// TIA Portal project "." (V14)

(* hardware
DEVICE "S7-1200 station_1"  S7-1200 Station
   slot 0: "Rack_0"  S7-1200 Rack  Rack  V1.0
   slot 1: "PLC_1"  CPU 1212C DC/DC/DC  6ES7 212-1AE31-0XB0  V3.0
   slot 2: "AI 4x13BIT/AQ 2x14BIT_1"  SM 1234 AI4/AQ2  6ES7 234-4HE30-0XB0  V1.0
   slot 3: "AI 4xRTD_1"  SM 1231 AI4 x RTD  6ES7 231-5PD32-0XB0  V2.0
   slot 101: "CM 1241 (RS485)_1"  CM 1241 (RS485)  6ES7 241-1CH30-0XB0  V1.0
DEVICE "HMI_1"  KTP600 Basic color PN
   slot 0: "KTP600 Basic color PN"  KTP600 Basic color PN  6AV6 647-0AD11-3AX0  12.0.0.0
   slot 1: "HMI_RT_1"  KTP600 Basic color PN  6AV6 647-0AD11-3AX0  12.0.0.0
   slot 5: "HMI_1.IE_CP_1"  PROFINET Interface  12.0.0.0
      slot 1: "Interfaz PROFINET_1"  PROFINET Interface
         slot 1: "Port_1"  Port
*)

// ===== PLC "PLC_1"  CPU 1212C DC/DC/DC =====

VAR_GLOBAL   // PLC tag table "Tabla de variables estándar"
   "Clock_10Hz" AT %M0.0 : Bool;
   "Clock_5Hz" AT %M0.1 : Bool;
   "Clock_2.5Hz" AT %M0.2 : Bool;
   "Clock_2Hz" AT %M0.3 : Bool;
   "Clock_1.25Hz" AT %M0.4 : Bool;
   "Clock_1Hz" AT %M0.5 : Bool;
   "Clock_0.625Hz" AT %M0.6 : Bool;
   "Clock_0.5Hz" AT %M0.7 : Bool;
   "ConexionExitosa" AT %M5.0 : Bool;
   "AlarmaDesconexion" AT %M5.1 : Bool;
   "A" AT %MW211 : Int;
   "System_Byte" AT %MB1 : Byte;
   "FirstScan" AT %M1.0 : Bool;
   "DiagStatusUpdate" AT %M1.1 : Bool;
   "AlwaysTRUE" AT %M1.2 : Bool;
   "AlwaysFALSE" AT %M1.3 : Bool;
   "ContadorAuxiliar" AT %MW200 : Int;
   "ModoManual" AT %M500.0 : Bool;
   "Tag_1" AT %MD66 : DWord;
   "Tag_2" AT %MD74 : DWord;
END_VAR

VAR_GLOBAL   // PLC tag table "Entradas y Salidas Fisicas"
   "Iniciar" AT %M800.1 : Bool;
   "Extraer" AT %M800.2 : Bool;
   "PilotoVerde" AT %Q0.0 : Bool;
   "PilotoAmarillo" AT %Q0.1 : Bool;
   "PilotoRojo" AT %Q0.2 : Bool;
   "IniciarbOTON" AT %I0.0 : Bool;
   "ExtraerBoton" AT %I0.1 : Bool;
END_VAR

VAR_GLOBAL   // PLC tag table "Memorias de Flanco"
   "Mem_Fer_FlancoBajadaIniciar" AT %M130.1 : Bool;
   "Mem_Fer_FlancoCompleta" AT %M130.2 : Bool;
   "Mem_Des_FlancoDestilado" AT %M131.0 : Bool;
   "Mem_Des_FlancoAgua" AT %M131.2 : Bool;
   "Mem_Rec_FlancoInicio" AT %M132.0 : Bool;
   "Mem_Rec_FlancoObjetivo" AT %M132.1 : Bool;
   "Mem_Rec_FlancoFin" AT %M132.2 : Bool;
   "AlertaAguaBajaDestilador" AT %M132.3 : Bool;
   "NivelBajoDestiador" AT %M132.4 : Bool;
   "Mem_ModoManual_Flanco" AT %M500.1 : Bool;
   "Pulso_SoltarActuadores" AT %M500.2 : Bool;
END_VAR

VAR_GLOBAL   // PLC tag table "Mediciones"
   "Fer_Temperatura" AT %MD40 : Real;
   "Des_Temperatura" AT %MD134 : Real;
   "Fer_Volumen" AT %MD54 : Real;
   "Des_Volumen" AT %MD14 : Real;
   "Rec_Volumen" AT %MD82 : Real;
   "RecirVol" AT %MD92 : Real;
END_VAR

VAR_GLOBAL   // PLC tag table "Estados"
   "Fer_FermentacionCompleta" AT %M72.7 : Bool;
   "Fer_Llenando" AT %M130.0 : Bool;
   "Des_CondicionesClarificar" AT %M131.1 : Bool;
   "AuxAlarmaFermentadorSobrecalentado" AT %MD158 : Real;
END_VAR

VAR_GLOBAL   // PLC tag table "Actuadores"
   "Act_BombaWash" AT %M36.0 : Bool;
   "Act_BombaAguaDestilador" AT %M36.1 : Bool;
   "Act_PurgaDestilador" AT %M36.2 : Bool;
   "Act_ValvRecirculadoDestilador" AT %M36.3 : Bool;
   "Act_ResistenciaDestilador" AT %M36.4 : Bool;
   "Act_ValvIngresoMosto" AT %M72.1 : Bool;
   "Act_PurgaFermentador" AT %M72.2 : Bool;
   "Act_RefrigeracionFermentador" AT %M72.5 : Bool;
   "Act_ValvVaciado" AT %M88.0 : Bool;
   "Act_BombaRecirculado" AT %M90.0 : Bool;
END_VAR

DATA_BLOCK "Proceso"   // DB1
{ S7_Optimized_Access := 'FALSE' }
VERSION : 0.1
   VAR
      Fer_VolInicialMosto : Real := 10.0;
      Fer_LimInfPerdida : Real := 8.12;
      Fer_LimSupTemp : Real := 20.5;
      Fer_LimInfTemp : Real := 19.5;
      Fer_UmbralSobrecalentado : Real := 22.125;
      Des_PesoInicialWash : Real := 0.0;
      Des_AguaAAgregar : Real := 0.0;
      Des_PesoFinal : Real := 0.0;
      Des_VolDescarteMetanol : Real := 0.0;
      Rec_VolBase : Real := 0.0;
      Rec_VolObjetivoRedestilado : Real := 0.0;
   END_VAR
BEGIN
END_DATA_BLOCK

DATA_BLOCK "DatosDeRecetas"   // DB4
{ S7_Optimized_Access := 'FALSE' }
VERSION : 0.1
   VAR
      NombreReceta : String := 'Irlandes';
      NombreReceta_1 : Int := 0;
      SetPointTempFermentador : Real := 20.0;
      HisterisisFermentador : Real := 0.5;
      SetPointTempDestilador : Real := 88.0;
      HisterisisDestilador : Real := 1.0;
      PorcAguaAgregada : Real := 15.0;
      PorcRedestilado : Real := 100.0;
      PorcPerdidaDescarte : Real := 6.125;
      PorcPerdidaFermentacion : Real := 4.0;
      PorcPurgaFermentador : Real := 10.0;
      PorcPurgaDestilador : Real := 5.0;
      CiclosRedestilado : Int := 2;
      VolumenPerdida : Real;
      Fer_LimInfVolumen : Real := 0.125;
      Fer_LimSupVolumen : Real := 52.125;
      Des_LimSupVolumen : Real := 50.125;
      Des_NivelBajo : Real := 0.2;
      Des_LimInfTemp : Real := 87.0;
      Des_LimSupTemp : Real := 89.125;
   END_VAR
BEGIN
END_DATA_BLOCK

DATA_BLOCK "Alarmas"   // DB6
{ S7_Optimized_Access := 'FALSE' }
VERSION : 0.1
   VAR
      Alm_FallaUSS : Bool;
      Alm_FermentadorSobrecalentado : Bool;
      Alm_AvisoDescarteMetanol : Bool;
      Alm_FermentadorLLeno : Bool;
      Alm_DemasiadoWashDestilador : Bool;
      Fase_MomentoDescarteMetanol : Bool;
      Fase_FermentacionTerminada : Bool;
      Fase_InicioLimpiezaFermentador : Bool;
      Fase_FinLimpiezaFermentador : Bool;
      Fase_InicioDestilado : Bool;
      Fase_InicioClarificado : Bool;
      Fase_DescarteExitoso : Bool;
      Fase_WhiskeyTerminado : Bool;
      Fase_InicioRecirculado : Bool;
      Fase_FinRecirculado : Bool;
      Fase_MezclaCompletada : Bool;
      Fase_ContadorRecirculado : Int;
      Vis_FinLimpiezaFermentador : Bool;
      Vis_InicioDestilado : Bool;
      Vis_DescarteExitoso : Bool;
      Vis_AvisoDescarteDeMetanol : Bool;
      aux1 : Bool;
      "aux 2" : Bool;
      AUx : Bool;
      Vis_FinRecirculado : Bool;
      Reserva_HMI : Bool;
   END_VAR
BEGIN
END_DATA_BLOCK

// folder: Control Manual

DATA_BLOCK "ControlManual"   // DB2
{ S7_Optimized_Access := 'FALSE' }
VERSION : 0.1
   VAR
      ManualBombaDeWash : Bool;
      ManualBombaDeAguaDestilador : Bool;
      ManualPurgaDestilador : Bool;
      ManualValvulaRecirculadoDestilador : Bool;
      ManualValvulaIngresoDeMosto : Bool;
      ManualPurgaFermentador : Bool;
      ManualEstadoRefriegeracionFermentador : Bool;
      ManualValvulaDeVaciado : Bool;
      ManualBombaDeRecirculado : Bool;
   END_VAR
BEGIN
END_DATA_BLOCK

// folder: System blocks/Program resources

DATA_BLOCK "IEC_Timer_0_DB"   // DB3
{ S7_Optimized_Access := 'TRUE' }
AUTHOR : Simatic
FAMILY : IEC
NAME : IEC_TMR
VERSION : 1.0
// stored: InstanceOfName IEC_TIMER
"IEC_TIMER"
BEGIN
END_DATA_BLOCK

DATA_BLOCK "IEC_Timer_0_DB_6"   // DB5
{ S7_Optimized_Access := 'TRUE' }
AUTHOR : Simatic
FAMILY : IEC
NAME : IEC_TMR
VERSION : 1.0
// stored: InstanceOfName IEC_TIMER
"IEC_TIMER"
BEGIN
END_DATA_BLOCK

DATA_BLOCK "IEC_Timer_0_DB_7"   // DB7
{ S7_Optimized_Access := 'TRUE' }
AUTHOR : Simatic
FAMILY : IEC
NAME : IEC_TMR
VERSION : 1.0
// stored: InstanceOfName IEC_TIMER
"IEC_TIMER"
BEGIN
END_DATA_BLOCK

DATA_BLOCK "IEC_Timer_0_DB_1"   // DB8
{ S7_Optimized_Access := 'TRUE' }
AUTHOR : Simatic
FAMILY : IEC
NAME : IEC_TMR
VERSION : 1.0
// stored: InstanceOfName IEC_TIMER
"IEC_TIMER"
BEGIN
END_DATA_BLOCK

DATA_BLOCK "IEC_Timer_0_DB_2"   // DB9
{ S7_Optimized_Access := 'TRUE' }
AUTHOR : Simatic
FAMILY : IEC
NAME : IEC_TMR
VERSION : 1.0
// stored: InstanceOfName IEC_TIMER
"IEC_TIMER"
BEGIN
END_DATA_BLOCK

DATA_BLOCK "IEC_Timer_0_DB_3"   // DB10
{ S7_Optimized_Access := 'TRUE' }
AUTHOR : Simatic
FAMILY : IEC
NAME : IEC_TMR
VERSION : 1.0
// stored: InstanceOfName IEC_TIMER
"IEC_TIMER"
BEGIN
END_DATA_BLOCK

DATA_BLOCK "IEC_Timer_0_DB_4"   // DB11
{ S7_Optimized_Access := 'TRUE' }
AUTHOR : Simatic
FAMILY : IEC
NAME : IEC_TMR
VERSION : 1.0
// stored: InstanceOfName IEC_TIMER
"IEC_TIMER"
BEGIN
END_DATA_BLOCK

DATA_BLOCK "IEC_Timer_0_DB_5"   // DB12
{ S7_Optimized_Access := 'TRUE' }
AUTHOR : Simatic
FAMILY : IEC
NAME : IEC_TMR
VERSION : 1.0
// stored: InstanceOfName IEC_TIMER
"IEC_TIMER"
BEGIN
END_DATA_BLOCK

DATA_BLOCK "IEC_Timer_0_DB_9"   // DB13
{ S7_Optimized_Access := 'TRUE' }
AUTHOR : Simatic
FAMILY : IEC
NAME : IEC_TMR
VERSION : 1.0
// stored: InstanceOfName IEC_TIMER
"IEC_TIMER"
BEGIN
END_DATA_BLOCK

DATA_BLOCK "IEC_Timer_0_DB_11"   // DB14
{ S7_Optimized_Access := 'TRUE' }
AUTHOR : Simatic
FAMILY : IEC
NAME : IEC_TMR
VERSION : 1.0
// stored: InstanceOfName IEC_TIMER
"IEC_TIMER"
BEGIN
END_DATA_BLOCK

DATA_BLOCK "IEC_Timer_0_DB_8"   // DB15
{ S7_Optimized_Access := 'TRUE' }
AUTHOR : Simatic
FAMILY : IEC
NAME : IEC_TMR
VERSION : 1.0
// stored: InstanceOfName IEC_TIMER
"IEC_TIMER"
BEGIN
END_DATA_BLOCK

DATA_BLOCK "IEC_Timer_0_DB_10"   // DB17
{ S7_Optimized_Access := 'TRUE' }
AUTHOR : Simatic
FAMILY : IEC
NAME : IEC_TMR
VERSION : 1.0
// stored: InstanceOfName IEC_TIMER
"IEC_TIMER"
BEGIN
END_DATA_BLOCK

// folder: (top level)

ORGANIZATION_BLOCK "control"   // OB126, LAD, ProgramCycle
TITLE = "Main Program Sweep (Cycle)"
{ S7_Optimized_Access := 'TRUE' }
VERSION : 0.1
   VAR_TEMP   // added for the SCL form of the ladder/FBD networks
      _w1 : Bool;
   END_VAR
BEGIN

REGION Network 1
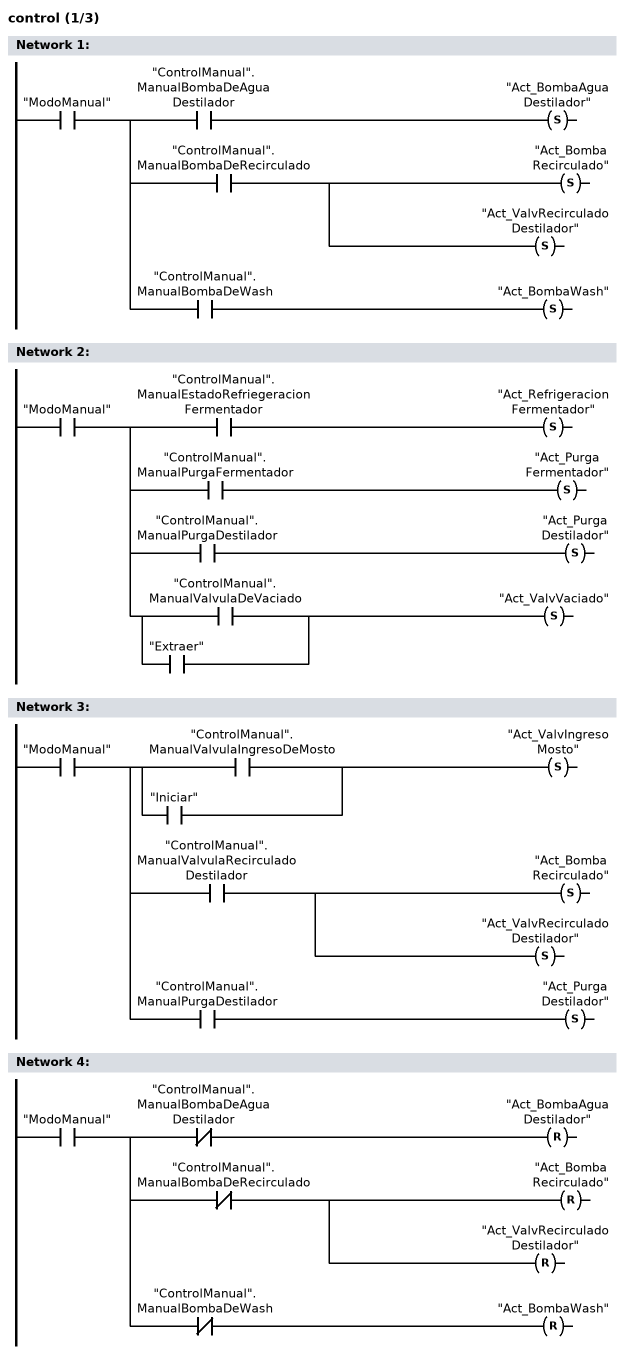
   RUNG wire#powerrail
      Contact( "ModoManual" )
      wire#w1
      Contact( "ControlManual".ManualBombaDeAguaDestilador )
      S_Coil( "Act_BombaAguaDestilador" )
   END_RUNG
   RUNG wire#w1
      Contact( "ControlManual".ManualBombaDeRecirculado )
      wire#w2
      S_Coil( "Act_BombaRecirculado" )
   END_RUNG
   RUNG wire#w2
      S_Coil( "Act_ValvRecirculadoDestilador" )
   END_RUNG
   RUNG wire#w1
      Contact( "ControlManual".ManualBombaDeWash )
      S_Coil( "Act_BombaWash" )
   END_RUNG
   // the same network as SCL:
   IF "ModoManual" AND "ControlManual".ManualBombaDeAguaDestilador THEN
       "Act_BombaAguaDestilador" := TRUE;
   END_IF;
   IF "ModoManual" AND "ControlManual".ManualBombaDeRecirculado THEN
       "Act_BombaRecirculado" := TRUE;
       "Act_ValvRecirculadoDestilador" := TRUE;
   END_IF;
   IF "ModoManual" AND "ControlManual".ManualBombaDeWash THEN "Act_BombaWash" := TRUE; END_IF;
END_REGION

REGION Network 2
   RUNG wire#powerrail
      Contact( "ModoManual" )
      wire#w1
      Contact( "ControlManual".ManualEstadoRefriegeracionFermentador )
      S_Coil( "Act_RefrigeracionFermentador" )
   END_RUNG
   RUNG wire#w1
      Contact( "ControlManual".ManualPurgaFermentador )
      S_Coil( "Act_PurgaFermentador" )
   END_RUNG
   RUNG wire#w1
      Contact( "ControlManual".ManualPurgaDestilador )
      S_Coil( "Act_PurgaDestilador" )
   END_RUNG
   RUNG wire#w1
      Contact( "ControlManual".ManualValvulaDeVaciado )
      wire#w2
      S_Coil( "Act_ValvVaciado" )
   END_RUNG
   RUNG wire#w1
      Contact( "Extraer" )
   END_RUNG wire#w2
   // the same network as SCL:
   IF "ModoManual" AND "ControlManual".ManualEstadoRefriegeracionFermentador THEN
       "Act_RefrigeracionFermentador" := TRUE;
   END_IF;
   IF "ModoManual" AND "ControlManual".ManualPurgaFermentador THEN "Act_PurgaFermentador" := TRUE; END_IF;
   IF "ModoManual" AND "ControlManual".ManualPurgaDestilador THEN "Act_PurgaDestilador" := TRUE; END_IF;
   IF "ModoManual" AND ("ControlManual".ManualValvulaDeVaciado OR "Extraer") THEN
       "Act_ValvVaciado" := TRUE;
   END_IF;
END_REGION

REGION Network 3
   RUNG wire#powerrail
      Contact( "ModoManual" )
      wire#w1
      Contact( "ControlManual".ManualValvulaIngresoDeMosto )
      wire#w2
      S_Coil( "Act_ValvIngresoMosto" )
   END_RUNG
   RUNG wire#w1
      Contact( "Iniciar" )
   END_RUNG wire#w2
   RUNG wire#w1
      Contact( "ControlManual".ManualValvulaRecirculadoDestilador )
      wire#w3
      S_Coil( "Act_BombaRecirculado" )
   END_RUNG
   RUNG wire#w3
      S_Coil( "Act_ValvRecirculadoDestilador" )
   END_RUNG
   RUNG wire#w1
      Contact( "ControlManual".ManualPurgaDestilador )
      S_Coil( "Act_PurgaDestilador" )
   END_RUNG
   // the same network as SCL:
   IF "ModoManual" AND ("ControlManual".ManualValvulaIngresoDeMosto OR "Iniciar") THEN
       "Act_ValvIngresoMosto" := TRUE;
   END_IF;
   IF "ModoManual" AND "ControlManual".ManualValvulaRecirculadoDestilador THEN
       "Act_BombaRecirculado" := TRUE;
       "Act_ValvRecirculadoDestilador" := TRUE;
   END_IF;
   IF "ModoManual" AND "ControlManual".ManualPurgaDestilador THEN "Act_PurgaDestilador" := TRUE; END_IF;
END_REGION

REGION Network 4
   RUNG wire#powerrail
      Contact( "ModoManual" )
      wire#w1
      I_Contact( "ControlManual".ManualBombaDeAguaDestilador )
      R_Coil( "Act_BombaAguaDestilador" )
   END_RUNG
   RUNG wire#w1
      I_Contact( "ControlManual".ManualBombaDeRecirculado )
      wire#w2
      R_Coil( "Act_BombaRecirculado" )
   END_RUNG
   RUNG wire#w2
      R_Coil( "Act_ValvRecirculadoDestilador" )
   END_RUNG
   RUNG wire#w1
      I_Contact( "ControlManual".ManualBombaDeWash )
      R_Coil( "Act_BombaWash" )
   END_RUNG
   // the same network as SCL:
   IF "ModoManual" AND NOT "ControlManual".ManualBombaDeAguaDestilador THEN
       "Act_BombaAguaDestilador" := FALSE;
   END_IF;
   IF "ModoManual" AND NOT "ControlManual".ManualBombaDeRecirculado THEN
       "Act_BombaRecirculado" := FALSE;
       "Act_ValvRecirculadoDestilador" := FALSE;
   END_IF;
   IF "ModoManual" AND NOT "ControlManual".ManualBombaDeWash THEN "Act_BombaWash" := FALSE; END_IF;
END_REGION

REGION Network 5
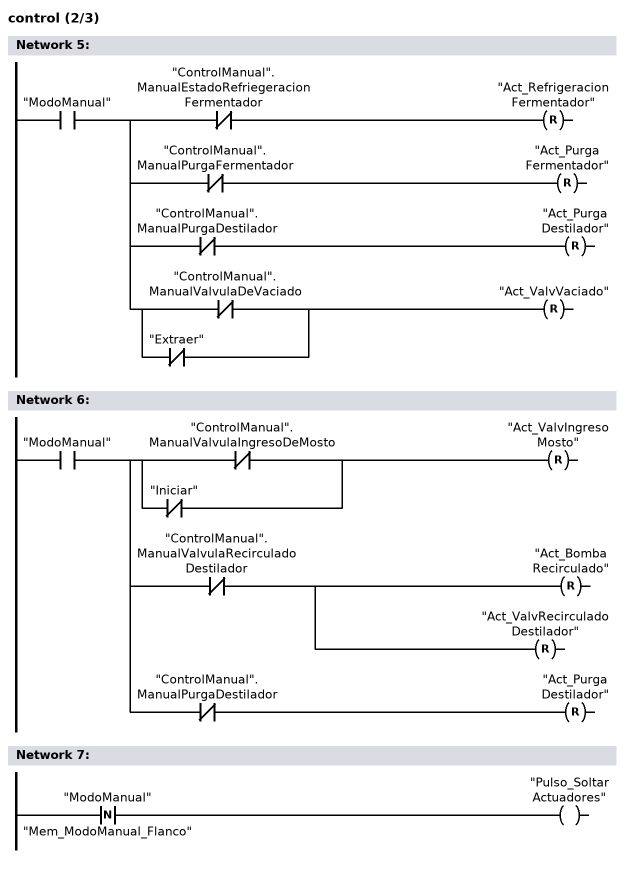
   RUNG wire#powerrail
      Contact( "ModoManual" )
      wire#w1
      I_Contact( "ControlManual".ManualEstadoRefriegeracionFermentador )
      R_Coil( "Act_RefrigeracionFermentador" )
   END_RUNG
   RUNG wire#w1
      I_Contact( "ControlManual".ManualPurgaFermentador )
      R_Coil( "Act_PurgaFermentador" )
   END_RUNG
   RUNG wire#w1
      I_Contact( "ControlManual".ManualPurgaDestilador )
      R_Coil( "Act_PurgaDestilador" )
   END_RUNG
   RUNG wire#w1
      I_Contact( "ControlManual".ManualValvulaDeVaciado )
      wire#w2
      R_Coil( "Act_ValvVaciado" )
   END_RUNG
   RUNG wire#w1
      I_Contact( "Extraer" )
   END_RUNG wire#w2
   // the same network as SCL:
   IF "ModoManual" AND NOT "ControlManual".ManualEstadoRefriegeracionFermentador THEN
       "Act_RefrigeracionFermentador" := FALSE;
   END_IF;
   IF "ModoManual" AND NOT "ControlManual".ManualPurgaFermentador THEN
       "Act_PurgaFermentador" := FALSE;
   END_IF;
   IF "ModoManual" AND NOT "ControlManual".ManualPurgaDestilador THEN "Act_PurgaDestilador" := FALSE; END_IF;
   IF "ModoManual" AND (NOT "ControlManual".ManualValvulaDeVaciado OR NOT "Extraer") THEN
       "Act_ValvVaciado" := FALSE;
   END_IF;
END_REGION

REGION Network 6
   RUNG wire#powerrail
      Contact( "ModoManual" )
      wire#w1
      I_Contact( "ControlManual".ManualValvulaIngresoDeMosto )
      wire#w2
      R_Coil( "Act_ValvIngresoMosto" )
   END_RUNG
   RUNG wire#w1
      I_Contact( "Iniciar" )
   END_RUNG wire#w2
   RUNG wire#w1
      I_Contact( "ControlManual".ManualValvulaRecirculadoDestilador )
      wire#w3
      R_Coil( "Act_BombaRecirculado" )
   END_RUNG
   RUNG wire#w3
      R_Coil( "Act_ValvRecirculadoDestilador" )
   END_RUNG
   RUNG wire#w1
      I_Contact( "ControlManual".ManualPurgaDestilador )
      R_Coil( "Act_PurgaDestilador" )
   END_RUNG
   // the same network as SCL:
   IF "ModoManual" AND (NOT "ControlManual".ManualValvulaIngresoDeMosto OR NOT "Iniciar") THEN
       "Act_ValvIngresoMosto" := FALSE;
   END_IF;
   IF "ModoManual" AND NOT "ControlManual".ManualValvulaRecirculadoDestilador THEN
       "Act_BombaRecirculado" := FALSE;
       "Act_ValvRecirculadoDestilador" := FALSE;
   END_IF;
   IF "ModoManual" AND NOT "ControlManual".ManualPurgaDestilador THEN "Act_PurgaDestilador" := FALSE; END_IF;
END_REGION

REGION Network 7
   RUNG wire#powerrail
      N_Contact(operand := "ModoManual", bit := "Mem_ModoManual_Flanco")
      Coil( "Pulso_SoltarActuadores" )
   END_RUNG
   // the same network as SCL:
   #_w1 := NOT "ModoManual" AND "Mem_ModoManual_Flanco";   // falling edge of "ModoManual"
   "Mem_ModoManual_Flanco" := "ModoManual";
   "Pulso_SoltarActuadores" := #_w1;
END_REGION

REGION Network 8
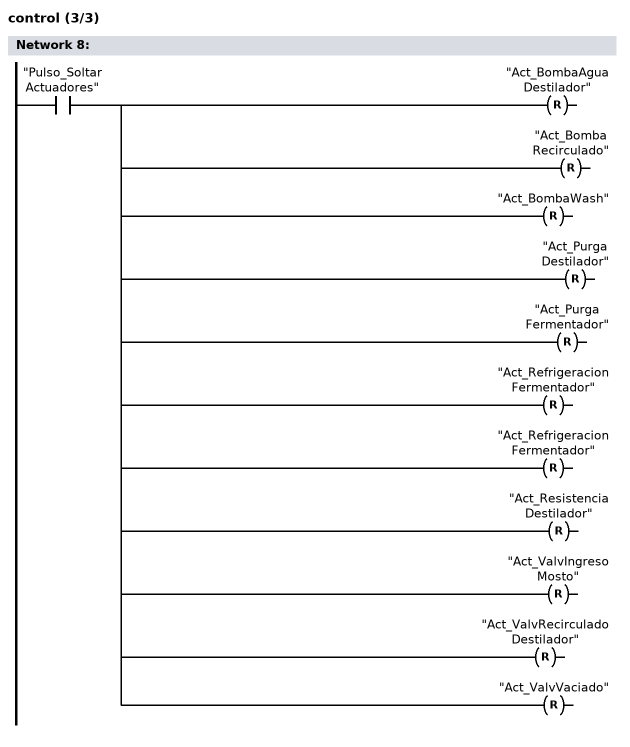
   RUNG wire#powerrail
      Contact( "Pulso_SoltarActuadores" )
      wire#w1
      R_Coil( "Act_BombaAguaDestilador" )
   END_RUNG
   RUNG wire#w1
      R_Coil( "Act_BombaRecirculado" )
   END_RUNG
   RUNG wire#w1
      R_Coil( "Act_BombaWash" )
   END_RUNG
   RUNG wire#w1
      R_Coil( "Act_PurgaDestilador" )
   END_RUNG
   RUNG wire#w1
      R_Coil( "Act_PurgaFermentador" )
   END_RUNG
   RUNG wire#w1
      R_Coil( "Act_RefrigeracionFermentador" )
   END_RUNG
   RUNG wire#w1
      R_Coil( "Act_RefrigeracionFermentador" )
   END_RUNG
   RUNG wire#w1
      R_Coil( "Act_ResistenciaDestilador" )
   END_RUNG
   RUNG wire#w1
      R_Coil( "Act_ValvIngresoMosto" )
   END_RUNG
   RUNG wire#w1
      R_Coil( "Act_ValvRecirculadoDestilador" )
   END_RUNG
   RUNG wire#w1
      R_Coil( "Act_ValvVaciado" )
   END_RUNG
   // the same network as SCL:
   IF "Pulso_SoltarActuadores" THEN
       "Act_BombaAguaDestilador" := FALSE;
       "Act_BombaRecirculado" := FALSE;
       "Act_BombaWash" := FALSE;
       "Act_PurgaDestilador" := FALSE;
       "Act_PurgaFermentador" := FALSE;
       "Act_RefrigeracionFermentador" := FALSE;
       "Act_RefrigeracionFermentador" := FALSE;
       "Act_ResistenciaDestilador" := FALSE;
       "Act_ValvIngresoMosto" := FALSE;
       "Act_ValvRecirculadoDestilador" := FALSE;
       "Act_ValvVaciado" := FALSE;
   END_IF;
END_REGION
END_ORGANIZATION_BLOCK

// folder: Control Manual

ORGANIZATION_BLOCK "Startup"   // OB100, LAD, Startup
TITLE = "Complete Restart"
{ S7_Optimized_Access := 'TRUE' }
VERSION : 0.1
   VAR_INPUT
      LostRetentive : Bool;   // True if retentive data are lost
      LostRTC : Bool;   // True if date and time are lost
   END_VAR
BEGIN

REGION Network 1
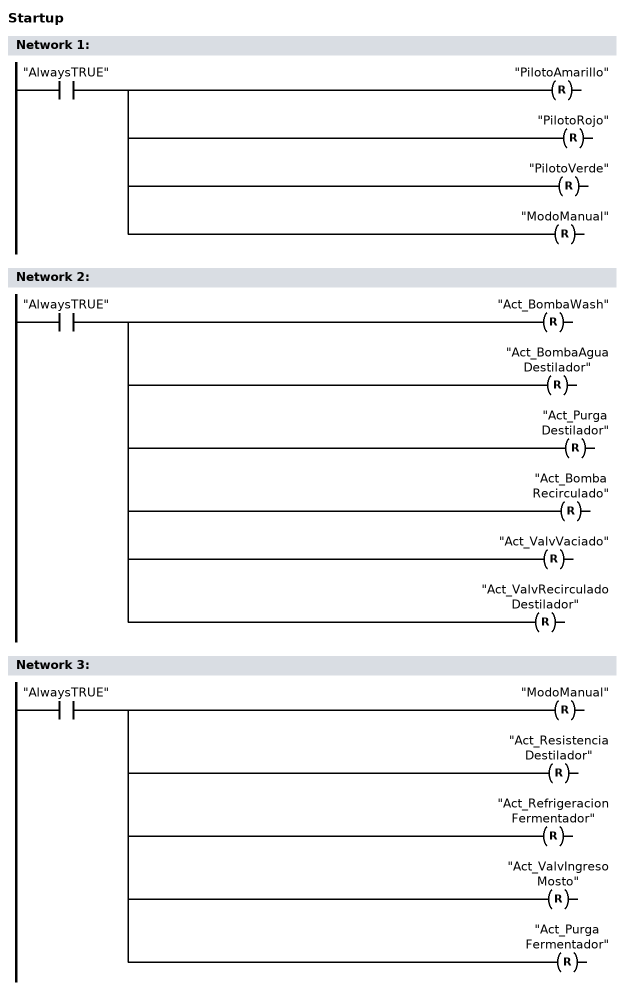
   RUNG wire#powerrail
      Contact( "AlwaysTRUE" )
      wire#w1
      R_Coil( "PilotoAmarillo" )
   END_RUNG
   RUNG wire#w1
      R_Coil( "PilotoRojo" )
   END_RUNG
   RUNG wire#w1
      R_Coil( "PilotoVerde" )
   END_RUNG
   RUNG wire#w1
      R_Coil( "ModoManual" )
   END_RUNG
   // the same network as SCL:
   IF "AlwaysTRUE" THEN
       "PilotoAmarillo" := FALSE;
       "PilotoRojo" := FALSE;
       "PilotoVerde" := FALSE;
       "ModoManual" := FALSE;
   END_IF;
END_REGION

REGION Network 2
   RUNG wire#powerrail
      Contact( "AlwaysTRUE" )
      wire#w1
      R_Coil( "Act_BombaWash" )
   END_RUNG
   RUNG wire#w1
      R_Coil( "Act_BombaAguaDestilador" )
   END_RUNG
   RUNG wire#w1
      R_Coil( "Act_PurgaDestilador" )
   END_RUNG
   RUNG wire#w1
      R_Coil( "Act_BombaRecirculado" )
   END_RUNG
   RUNG wire#w1
      R_Coil( "Act_ValvVaciado" )
   END_RUNG
   RUNG wire#w1
      R_Coil( "Act_ValvRecirculadoDestilador" )
   END_RUNG
   // the same network as SCL:
   IF "AlwaysTRUE" THEN
       "Act_BombaWash" := FALSE;
       "Act_BombaAguaDestilador" := FALSE;
       "Act_PurgaDestilador" := FALSE;
       "Act_BombaRecirculado" := FALSE;
       "Act_ValvVaciado" := FALSE;
       "Act_ValvRecirculadoDestilador" := FALSE;
   END_IF;
END_REGION

REGION Network 3
   RUNG wire#powerrail
      Contact( "AlwaysTRUE" )
      wire#w1
      R_Coil( "ModoManual" )
   END_RUNG
   RUNG wire#w1
      R_Coil( "Act_ResistenciaDestilador" )
   END_RUNG
   RUNG wire#w1
      R_Coil( "Act_RefrigeracionFermentador" )
   END_RUNG
   RUNG wire#w1
      R_Coil( "Act_ValvIngresoMosto" )
   END_RUNG
   RUNG wire#w1
      R_Coil( "Act_PurgaFermentador" )
   END_RUNG
   // the same network as SCL:
   IF "AlwaysTRUE" THEN
       "ModoManual" := FALSE;
       "Act_ResistenciaDestilador" := FALSE;
       "Act_RefrigeracionFermentador" := FALSE;
       "Act_ValvIngresoMosto" := FALSE;
       "Act_PurgaFermentador" := FALSE;
   END_IF;
END_REGION
END_ORGANIZATION_BLOCK

// folder: Destilador

ORGANIZATION_BLOCK "Control de Temperatura destilador"   // OB31, LAD, CyclicInterrupt
{ S7_Optimized_Access := 'TRUE' }
VERSION : 0.1
   VAR_TEMP   // added for the SCL form of the ladder/FBD networks
      _w1 : Bool;
      _w2 : Bool;
   END_VAR
BEGIN

REGION Network 1: Control
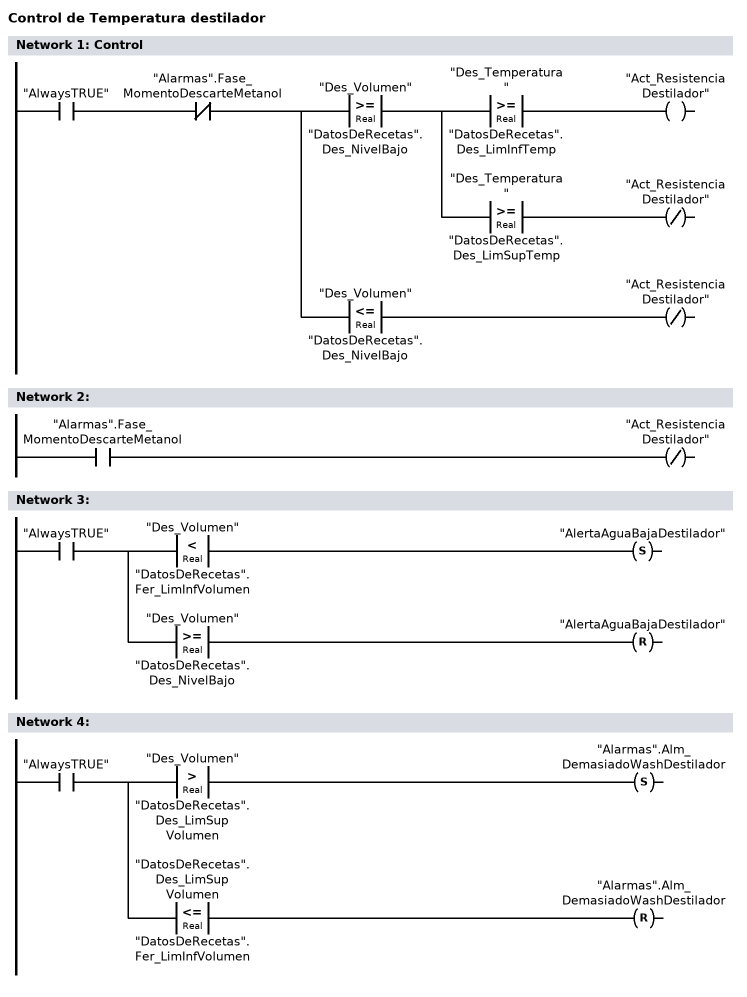
   RUNG wire#powerrail
      Contact( "AlwaysTRUE" )
      I_Contact( "Alarmas".Fase_MomentoDescarteMetanol )
      wire#w1
      { S7_Templates := "SrcType := Real" } GE_Contact(in1 := "Des_Volumen", in2 := "DatosDeRecetas".Des_NivelBajo)
      wire#w2
      { S7_Templates := "SrcType := Real" } GE_Contact(in1 := "Des_Temperatura", in2 := "DatosDeRecetas".Des_LimInfTemp)
      Coil( "Act_ResistenciaDestilador" )
   END_RUNG
   RUNG wire#w2
      { S7_Templates := "SrcType := Real" } GE_Contact(in1 := "Des_Temperatura", in2 := "DatosDeRecetas".Des_LimSupTemp)
      I_Coil( "Act_ResistenciaDestilador" )
   END_RUNG
   RUNG wire#w1
      { S7_Templates := "SrcType := Real" } LE_Contact(in1 := "Des_Volumen", in2 := "DatosDeRecetas".Des_NivelBajo)
      I_Coil( "Act_ResistenciaDestilador" )
   END_RUNG
   // the same network as SCL:
   #_w1 := "AlwaysTRUE" AND NOT "Alarmas".Fase_MomentoDescarteMetanol;
   #_w2 := #_w1 AND ("Des_Volumen" >= "DatosDeRecetas".Des_NivelBajo);
   "Act_ResistenciaDestilador" := #_w2 AND ("Des_Temperatura" >= "DatosDeRecetas".Des_LimInfTemp);
   "Act_ResistenciaDestilador" := NOT (#_w2 AND ("Des_Temperatura" >= "DatosDeRecetas".Des_LimSupTemp));
   "Act_ResistenciaDestilador" := NOT (#_w1 AND ("Des_Volumen" <= "DatosDeRecetas".Des_NivelBajo));
END_REGION

REGION Network 2
   RUNG wire#powerrail
      Contact( "Alarmas".Fase_MomentoDescarteMetanol )
      I_Coil( "Act_ResistenciaDestilador" )
   END_RUNG
   // the same network as SCL:
   "Act_ResistenciaDestilador" := NOT "Alarmas".Fase_MomentoDescarteMetanol;
END_REGION

REGION Network 3
   RUNG wire#powerrail
      Contact( "AlwaysTRUE" )
      wire#w1
      { S7_Templates := "SrcType := Real" } LT_Contact(in1 := "Des_Volumen", in2 := "DatosDeRecetas".Fer_LimInfVolumen)
      S_Coil( "AlertaAguaBajaDestilador" )
   END_RUNG
   RUNG wire#w1
      { S7_Templates := "SrcType := Real" } GE_Contact(in1 := "Des_Volumen", in2 := "DatosDeRecetas".Des_NivelBajo)
      R_Coil( "AlertaAguaBajaDestilador" )
   END_RUNG
   // the same network as SCL:
   IF "AlwaysTRUE" AND ("Des_Volumen" < "DatosDeRecetas".Fer_LimInfVolumen) THEN
       "AlertaAguaBajaDestilador" := TRUE;
   END_IF;
   IF "AlwaysTRUE" AND ("Des_Volumen" >= "DatosDeRecetas".Des_NivelBajo) THEN
       "AlertaAguaBajaDestilador" := FALSE;
   END_IF;
END_REGION

REGION Network 4
   RUNG wire#powerrail
      Contact( "AlwaysTRUE" )
      wire#w1
      { S7_Templates := "SrcType := Real" } GT_Contact(in1 := "Des_Volumen", in2 := "DatosDeRecetas".Des_LimSupVolumen)
      S_Coil( "Alarmas".Alm_DemasiadoWashDestilador )
   END_RUNG
   RUNG wire#w1
      { S7_Templates := "SrcType := Real" } LE_Contact(in1 := "DatosDeRecetas".Des_LimSupVolumen, in2 := "DatosDeRecetas".Fer_LimInfVolumen)
      R_Coil( "Alarmas".Alm_DemasiadoWashDestilador )
   END_RUNG
   // the same network as SCL:
   IF "AlwaysTRUE" AND ("Des_Volumen" > "DatosDeRecetas".Des_LimSupVolumen) THEN
       "Alarmas".Alm_DemasiadoWashDestilador := TRUE;
   END_IF;
   IF "AlwaysTRUE" AND ("DatosDeRecetas".Des_LimSupVolumen <= "DatosDeRecetas".Fer_LimInfVolumen) THEN
       "Alarmas".Alm_DemasiadoWashDestilador := FALSE;
   END_IF;
END_REGION
END_ORGANIZATION_BLOCK

ORGANIZATION_BLOCK "Configuracion y ciclo de programa"   // OB124, LAD, ProgramCycle
TITLE = "Main Program Sweep (Cycle)"
{ S7_Optimized_Access := 'TRUE' }
VERSION : 0.1
   VAR_TEMP
      PesoInicialDelWash : Real;
      Temp_1 : Bool;
      PesoFinal : Real;
      AguaAAgregar : Real;
      PesoDeMetanol : Real;
   END_VAR
   VAR_TEMP   // added for the SCL form of the ladder/FBD networks
      _w1 : Bool;
   END_VAR
BEGIN

REGION Network 1: Pesaje previo al clarificado
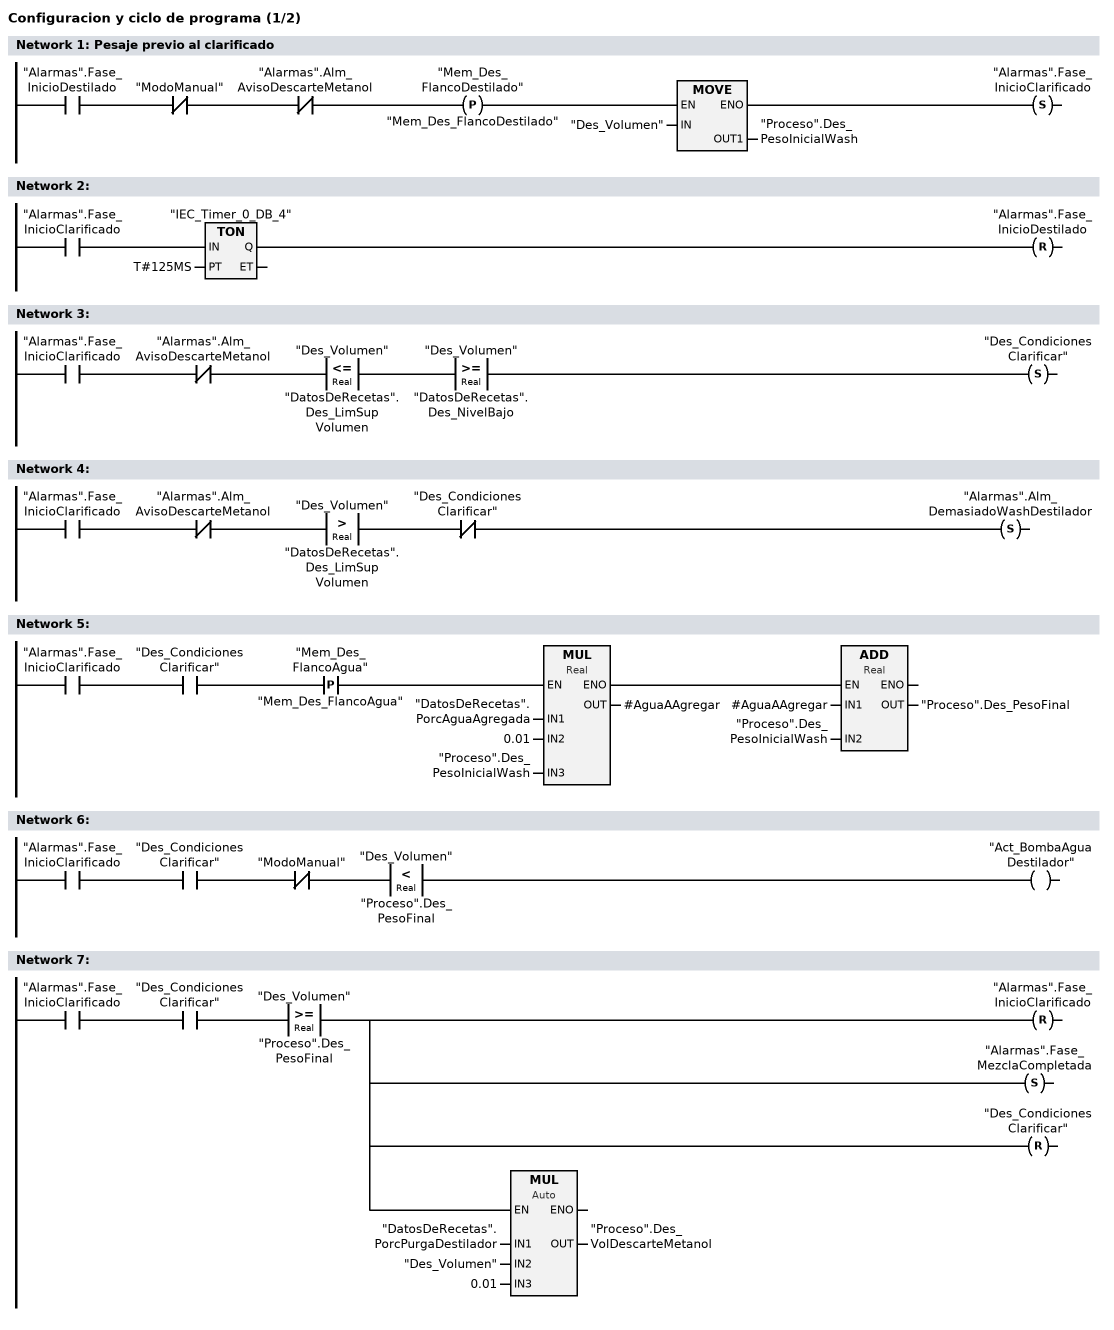
   // ENO of a box is taken as its EN; it also drops when the box reports an error
   #_w1 := "Alarmas".Fase_InicioDestilado AND NOT "ModoManual" AND NOT "Alarmas".Alm_AvisoDescarteMetanol;
   "Mem_Des_FlancoDestilado" := #_w1 AND NOT "Mem_Des_FlancoDestilado";   // rising edge
   "Mem_Des_FlancoDestilado" := #_w1;
   IF #_w1 THEN
       "Proceso".Des_PesoInicialWash := "Des_Volumen";
       "Alarmas".Fase_InicioClarificado := TRUE;
   END_IF;
END_REGION

REGION Network 2
   "IEC_Timer_0_DB_4".TON(IN := "Alarmas".Fase_InicioClarificado, PT := T#125MS);
   IF "IEC_Timer_0_DB_4".Q THEN "Alarmas".Fase_InicioDestilado := FALSE; END_IF;
END_REGION

REGION Network 3
   RUNG wire#powerrail
      Contact( "Alarmas".Fase_InicioClarificado )
      I_Contact( "Alarmas".Alm_AvisoDescarteMetanol )
      { S7_Templates := "SrcType := Real" } LE_Contact(in1 := "Des_Volumen", in2 := "DatosDeRecetas".Des_LimSupVolumen)
      { S7_Templates := "SrcType := Real" } GE_Contact(in1 := "Des_Volumen", in2 := "DatosDeRecetas".Des_NivelBajo)
      S_Coil( "Des_CondicionesClarificar" )
   END_RUNG
   // the same network as SCL:
   IF "Alarmas".Fase_InicioClarificado AND NOT "Alarmas".Alm_AvisoDescarteMetanol AND ("Des_Volumen" <= "DatosDeRecetas".Des_LimSupVolumen) AND ("Des_Volumen" >= "DatosDeRecetas".Des_NivelBajo) THEN
       "Des_CondicionesClarificar" := TRUE;
   END_IF;
END_REGION

REGION Network 4
   RUNG wire#powerrail
      Contact( "Alarmas".Fase_InicioClarificado )
      I_Contact( "Alarmas".Alm_AvisoDescarteMetanol )
      { S7_Templates := "SrcType := Real" } GT_Contact(in1 := "Des_Volumen", in2 := "DatosDeRecetas".Des_LimSupVolumen)
      I_Contact( "Des_CondicionesClarificar" )
      S_Coil( "Alarmas".Alm_DemasiadoWashDestilador )
   END_RUNG
   // the same network as SCL:
   IF "Alarmas".Fase_InicioClarificado AND NOT "Alarmas".Alm_AvisoDescarteMetanol AND ("Des_Volumen" > "DatosDeRecetas".Des_LimSupVolumen) AND NOT "Des_CondicionesClarificar" THEN
       "Alarmas".Alm_DemasiadoWashDestilador := TRUE;
   END_IF;
END_REGION

REGION Network 5
   RUNG wire#powerrail
      Contact( "Alarmas".Fase_InicioClarificado )
      Contact( "Des_CondicionesClarificar" )
      P_Contact(operand := "Mem_Des_FlancoAgua", bit := "Mem_Des_FlancoAgua")
      { S7_Templates := "SrcType := Real"; S7_GenerateENO := "TRUE" } Mul(in1 := "DatosDeRecetas".PorcAguaAgregada, in2 := 0.01, in3 := "Proceso".Des_PesoInicialWash, out => #AguaAAgregar)
      { S7_Templates := "SrcType := Real"; S7_GenerateENO := "TRUE" } Add(in1 := #AguaAAgregar, in2 := "Proceso".Des_PesoInicialWash, out => "Proceso".Des_PesoFinal)
   END_RUNG
   // the same network as SCL:
   // ENO of a box is taken as its EN; it also drops when the box reports an error
   #_w1 := "Alarmas".Fase_InicioClarificado AND "Des_CondicionesClarificar" AND "Mem_Des_FlancoAgua" AND NOT "Mem_Des_FlancoAgua";   // rising edge of "Mem_Des_FlancoAgua"
   "Mem_Des_FlancoAgua" := "Mem_Des_FlancoAgua";
   IF #_w1 THEN
       #AguaAAgregar := "DatosDeRecetas".PorcAguaAgregada * 0.01 * "Proceso".Des_PesoInicialWash;
       "Proceso".Des_PesoFinal := #AguaAAgregar + "Proceso".Des_PesoInicialWash;
   END_IF;
END_REGION

REGION Network 6
   RUNG wire#powerrail
      Contact( "Alarmas".Fase_InicioClarificado )
      Contact( "Des_CondicionesClarificar" )
      I_Contact( "ModoManual" )
      { S7_Templates := "SrcType := Real" } LT_Contact(in1 := "Des_Volumen", in2 := "Proceso".Des_PesoFinal)
      Coil( "Act_BombaAguaDestilador" )
   END_RUNG
   // the same network as SCL:
   "Act_BombaAguaDestilador" := "Alarmas".Fase_InicioClarificado AND "Des_CondicionesClarificar" AND NOT "ModoManual" AND ("Des_Volumen" < "Proceso".Des_PesoFinal);
END_REGION

REGION Network 7
   RUNG wire#powerrail
      Contact( "Alarmas".Fase_InicioClarificado )
      Contact( "Des_CondicionesClarificar" )
      { S7_Templates := "SrcType := Real" } GE_Contact(in1 := "Des_Volumen", in2 := "Proceso".Des_PesoFinal)
      wire#w1
      R_Coil( "Alarmas".Fase_InicioClarificado )
   END_RUNG
   RUNG wire#w1
      S_Coil( "Alarmas".Fase_MezclaCompletada )
   END_RUNG
   RUNG wire#w1
      R_Coil( "Des_CondicionesClarificar" )
   END_RUNG
   RUNG wire#w1
      { S7_GenerateENO := "TRUE" } Mul(in1 := "DatosDeRecetas".PorcPurgaDestilador, in2 := "Des_Volumen", in3 := 0.01, out => "Proceso".Des_VolDescarteMetanol)
   END_RUNG
   // the same network as SCL:
   #_w1 := "Alarmas".Fase_InicioClarificado AND "Des_CondicionesClarificar" AND ("Des_Volumen" >= "Proceso".Des_PesoFinal);
   IF #_w1 THEN
       "Alarmas".Fase_InicioClarificado := FALSE;
       "Alarmas".Fase_MezclaCompletada := TRUE;
       "Des_CondicionesClarificar" := FALSE;
       "Proceso".Des_VolDescarteMetanol := "DatosDeRecetas".PorcPurgaDestilador * "Des_Volumen" * 0.01;
   END_IF;
END_REGION

REGION Network 8
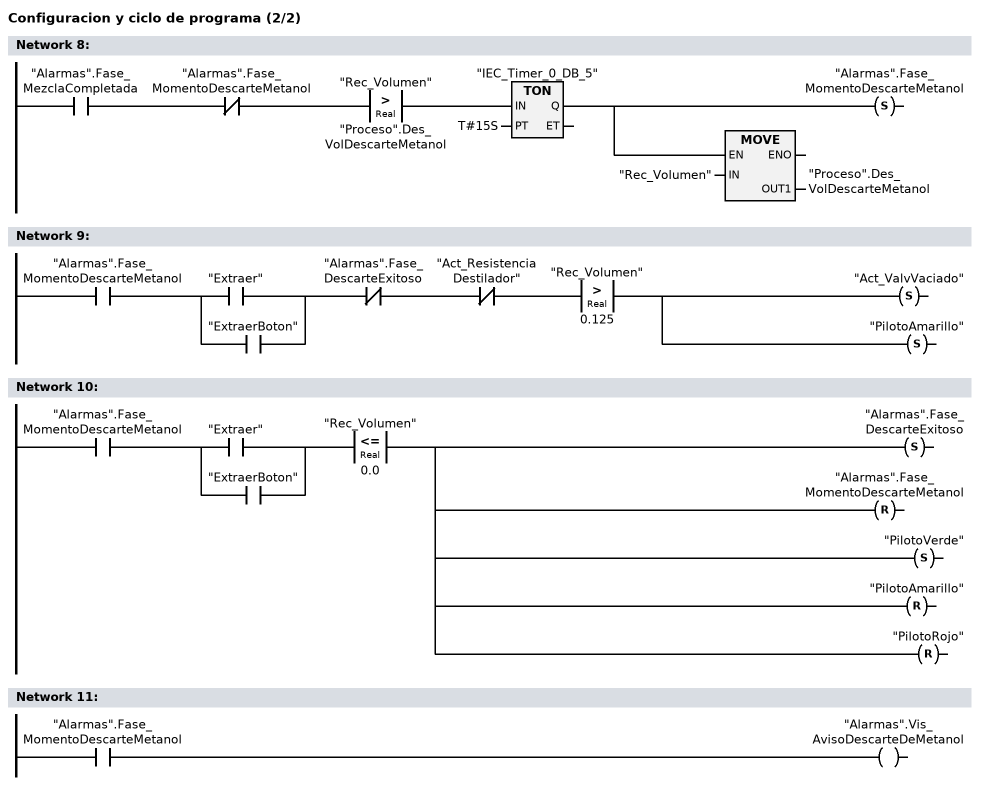
   "IEC_Timer_0_DB_5".TON(IN := "Alarmas".Fase_MezclaCompletada AND NOT "Alarmas".Fase_MomentoDescarteMetanol AND ("Rec_Volumen" > "Proceso".Des_VolDescarteMetanol),
                          PT := T#15S);
   IF "IEC_Timer_0_DB_5".Q THEN
       "Alarmas".Fase_MomentoDescarteMetanol := TRUE;
       "Proceso".Des_VolDescarteMetanol := "Rec_Volumen";
   END_IF;
END_REGION

REGION Network 9
   RUNG wire#powerrail
      Contact( "Alarmas".Fase_MomentoDescarteMetanol )
      wire#w1
      Contact( "Extraer" )
      wire#w2
      I_Contact( "Alarmas".Fase_DescarteExitoso )
      I_Contact( "Act_ResistenciaDestilador" )
      { S7_Templates := "SrcType := Real" } GT_Contact(in1 := "Rec_Volumen", in2 := 0.125)
      wire#w3
      S_Coil( "Act_ValvVaciado" )
   END_RUNG
   RUNG wire#w1
      Contact( "ExtraerBoton" )
   END_RUNG wire#w2
   RUNG wire#w3
      S_Coil( "PilotoAmarillo" )
   END_RUNG
   // the same network as SCL:
   IF "Alarmas".Fase_MomentoDescarteMetanol AND ("Extraer" OR "ExtraerBoton") AND NOT "Alarmas".Fase_DescarteExitoso AND NOT "Act_ResistenciaDestilador" AND ("Rec_Volumen" > 0.125) THEN
       "Act_ValvVaciado" := TRUE;
       "PilotoAmarillo" := TRUE;
   END_IF;
END_REGION

REGION Network 10
   RUNG wire#powerrail
      Contact( "Alarmas".Fase_MomentoDescarteMetanol )
      wire#w1
      Contact( "Extraer" )
      wire#w2
      { S7_Templates := "SrcType := Real" } LE_Contact(in1 := "Rec_Volumen", in2 := 0.0)
      wire#w3
      S_Coil( "Alarmas".Fase_DescarteExitoso )
   END_RUNG
   RUNG wire#w1
      Contact( "ExtraerBoton" )
   END_RUNG wire#w2
   RUNG wire#w3
      R_Coil( "Alarmas".Fase_MomentoDescarteMetanol )
   END_RUNG
   RUNG wire#w3
      S_Coil( "PilotoVerde" )
   END_RUNG
   RUNG wire#w3
      R_Coil( "PilotoAmarillo" )
   END_RUNG
   RUNG wire#w3
      R_Coil( "PilotoRojo" )
   END_RUNG
   // the same network as SCL:
   IF "Alarmas".Fase_MomentoDescarteMetanol AND ("Extraer" OR "ExtraerBoton") AND ("Rec_Volumen" <= 0.0) THEN
       "Alarmas".Fase_DescarteExitoso := TRUE;
   END_IF;
   #_w1 := "Alarmas".Fase_MomentoDescarteMetanol AND ("Extraer" OR "ExtraerBoton") AND ("Rec_Volumen" <= 0.0);
   IF #_w1 THEN
       "Alarmas".Fase_MomentoDescarteMetanol := FALSE;
       "PilotoVerde" := TRUE;
       "PilotoAmarillo" := FALSE;
       "PilotoRojo" := FALSE;
   END_IF;
END_REGION

REGION Network 11
   RUNG wire#powerrail
      Contact( "Alarmas".Fase_MomentoDescarteMetanol )
      Coil( "Alarmas".Vis_AvisoDescarteDeMetanol )
   END_RUNG
   // the same network as SCL:
   "Alarmas".Vis_AvisoDescarteDeMetanol := "Alarmas".Fase_MomentoDescarteMetanol;
END_REGION
END_ORGANIZATION_BLOCK

ORGANIZATION_BLOCK "Calcular  limites on off destilador"   // OB127, LAD, ProgramCycle
TITLE = "Main Program Sweep (Cycle)"
{ S7_Optimized_Access := 'TRUE' }
VERSION : 0.1
BEGIN

REGION Network 1
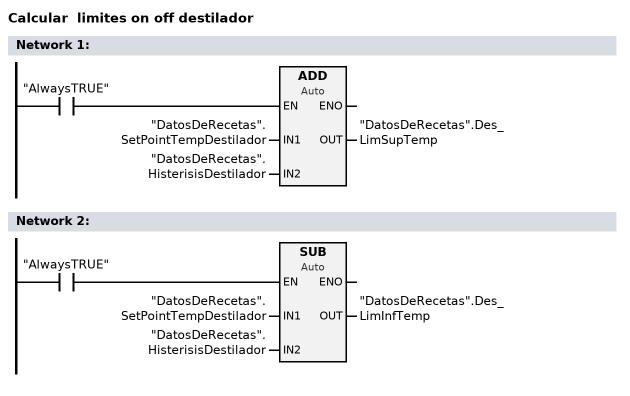
   RUNG wire#powerrail
      Contact( "AlwaysTRUE" )
      { S7_GenerateENO := "TRUE" } Add(in1 := "DatosDeRecetas".SetPointTempDestilador, in2 := "DatosDeRecetas".HisterisisDestilador, out => "DatosDeRecetas".Des_LimSupTemp)
   END_RUNG
   // the same network as SCL:
   IF "AlwaysTRUE" THEN
       "DatosDeRecetas".Des_LimSupTemp := "DatosDeRecetas".SetPointTempDestilador + "DatosDeRecetas".HisterisisDestilador;
   END_IF;
END_REGION

REGION Network 2
   RUNG wire#powerrail
      Contact( "AlwaysTRUE" )
      { S7_GenerateENO := "TRUE" } Sub(in1 := "DatosDeRecetas".SetPointTempDestilador, in2 := "DatosDeRecetas".HisterisisDestilador, out => "DatosDeRecetas".Des_LimInfTemp)
   END_RUNG
   // the same network as SCL:
   IF "AlwaysTRUE" THEN
       "DatosDeRecetas".Des_LimInfTemp := "DatosDeRecetas".SetPointTempDestilador - "DatosDeRecetas".HisterisisDestilador;
   END_IF;
END_REGION
END_ORGANIZATION_BLOCK

// folder: Fermentador

ORGANIZATION_BLOCK "Control de ingreso Mosto y salida de Wash"   // OB1, LAD, ProgramCycle
TITLE = "Control del Mosto y Wash Fermentador"
{ S7_Optimized_Access := 'TRUE' }
VERSION : 0.1
   VAR_TEMP
      Auxiliarrr : Real;
      FlancoDeBajadaInicio : Bool;
      Temp_1 : Bool;
      Auxiliar : Bool;
   END_VAR
   VAR_TEMP   // added for the SCL form of the ladder/FBD networks
      _w1 : Bool;
   END_VAR
BEGIN

REGION Network 1
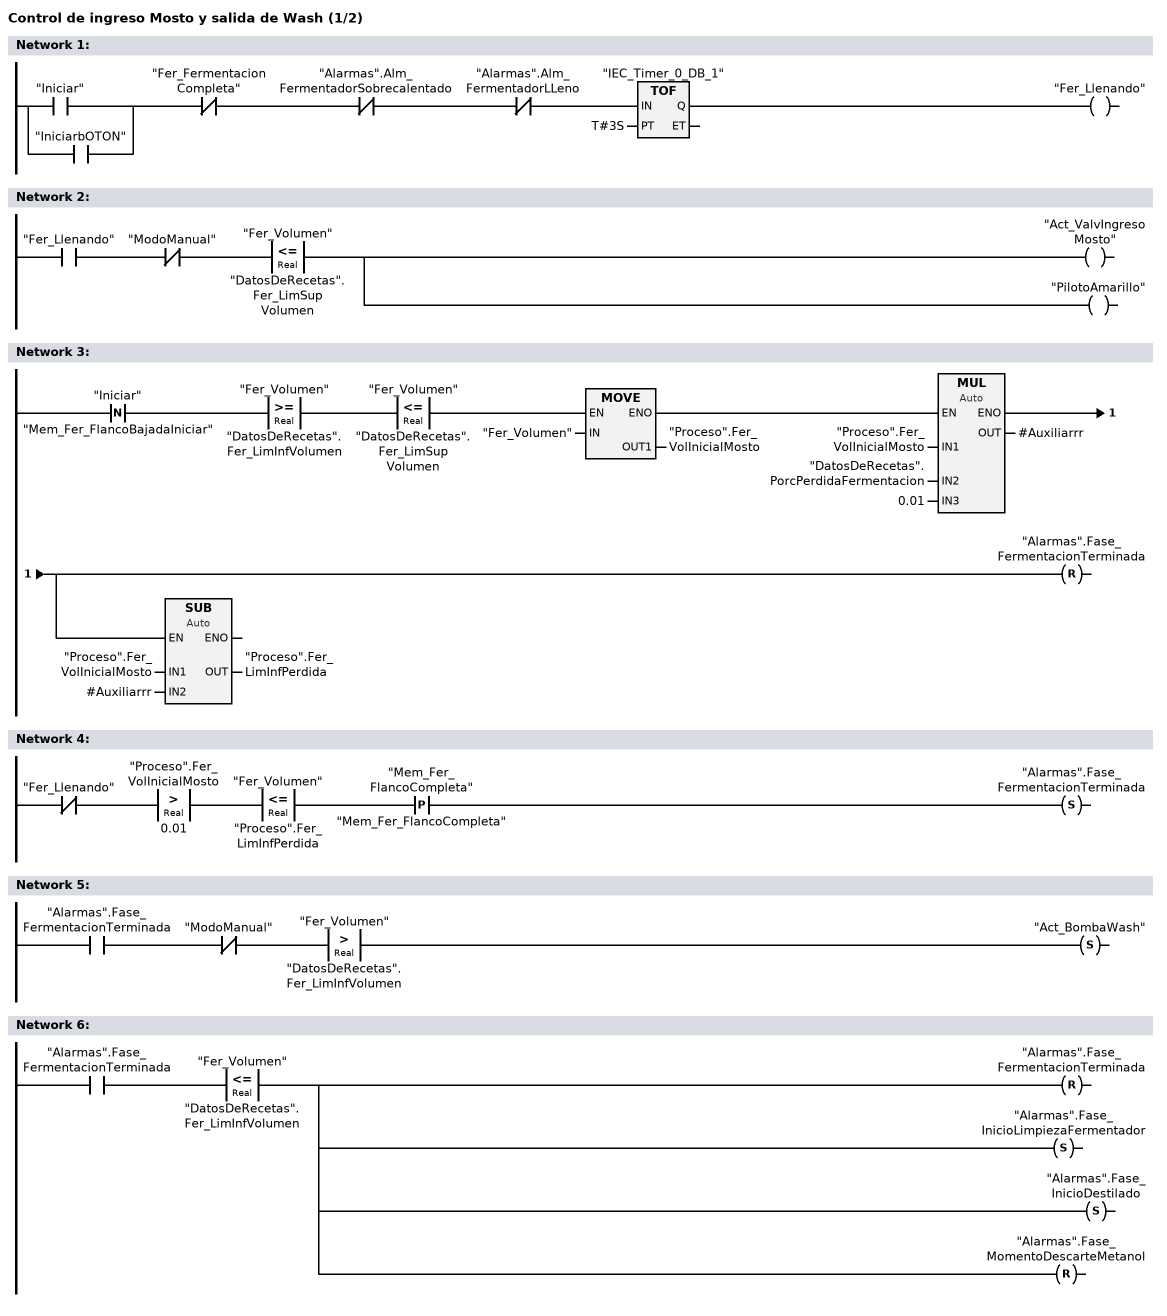
   "IEC_Timer_0_DB_1".TOF(IN := ("Iniciar" OR "IniciarbOTON") AND NOT "Fer_FermentacionCompleta" AND NOT "Alarmas".Alm_FermentadorSobrecalentado AND NOT "Alarmas".Alm_FermentadorLLeno,
                          PT := T#3S);
   "Fer_Llenando" := "IEC_Timer_0_DB_1".Q;
END_REGION

REGION Network 2
   RUNG wire#powerrail
      Contact( "Fer_Llenando" )
      I_Contact( "ModoManual" )
      { S7_Templates := "SrcType := Real" } LE_Contact(in1 := "Fer_Volumen", in2 := "DatosDeRecetas".Fer_LimSupVolumen)
      wire#w1
      Coil( "Act_ValvIngresoMosto" )
   END_RUNG
   RUNG wire#w1
      Coil( "PilotoAmarillo" )
   END_RUNG
   // the same network as SCL:
   "Act_ValvIngresoMosto" := "Fer_Llenando" AND NOT "ModoManual" AND ("Fer_Volumen" <= "DatosDeRecetas".Fer_LimSupVolumen);
   "PilotoAmarillo" := "Act_ValvIngresoMosto";
END_REGION

REGION Network 3
   RUNG wire#powerrail
      N_Contact(operand := "Iniciar", bit := "Mem_Fer_FlancoBajadaIniciar")
      { S7_Templates := "SrcType := Real" } GE_Contact(in1 := "Fer_Volumen", in2 := "DatosDeRecetas".Fer_LimInfVolumen)
      { S7_Templates := "SrcType := Real" } LE_Contact(in1 := "Fer_Volumen", in2 := "DatosDeRecetas".Fer_LimSupVolumen)
      { S7_GenerateENO := "TRUE" } Move(in := "Fer_Volumen", out1 => "Proceso".Fer_VolInicialMosto)
      { S7_GenerateENO := "TRUE" } Mul(in1 := "Proceso".Fer_VolInicialMosto, in2 := "DatosDeRecetas".PorcPerdidaFermentacion, in3 := 0.01, out => #Auxiliarrr)
      wire#w1
      R_Coil( "Alarmas".Fase_FermentacionTerminada )
   END_RUNG
   RUNG wire#w1
      { S7_GenerateENO := "TRUE" } Sub(in1 := "Proceso".Fer_VolInicialMosto, in2 := #Auxiliarrr, out => "Proceso".Fer_LimInfPerdida)
   END_RUNG
   // the same network as SCL:
   // ENO of a box is taken as its EN; it also drops when the box reports an error
   #_w1 := NOT "Iniciar" AND "Mem_Fer_FlancoBajadaIniciar";   // falling edge of "Iniciar"
   "Mem_Fer_FlancoBajadaIniciar" := "Iniciar";
   IF #_w1 AND ("Fer_Volumen" >= "DatosDeRecetas".Fer_LimInfVolumen) AND ("Fer_Volumen" <= "DatosDeRecetas".Fer_LimSupVolumen) THEN
       "Proceso".Fer_VolInicialMosto := "Fer_Volumen";
       #Auxiliarrr := "Proceso".Fer_VolInicialMosto * "DatosDeRecetas".PorcPerdidaFermentacion * 0.01;
       "Alarmas".Fase_FermentacionTerminada := FALSE;
       "Proceso".Fer_LimInfPerdida := "Proceso".Fer_VolInicialMosto - #Auxiliarrr;
   END_IF;
END_REGION

REGION Network 4
   RUNG wire#powerrail
      I_Contact( "Fer_Llenando" )
      { S7_Templates := "SrcType := Real" } GT_Contact(in1 := "Proceso".Fer_VolInicialMosto, in2 := 0.01)
      { S7_Templates := "SrcType := Real" } LE_Contact(in1 := "Fer_Volumen", in2 := "Proceso".Fer_LimInfPerdida)
      P_Contact(operand := "Mem_Fer_FlancoCompleta", bit := "Mem_Fer_FlancoCompleta")
      S_Coil( "Alarmas".Fase_FermentacionTerminada )
   END_RUNG
   // the same network as SCL:
   #_w1 := NOT "Fer_Llenando" AND ("Proceso".Fer_VolInicialMosto > 0.01) AND ("Fer_Volumen" <= "Proceso".Fer_LimInfPerdida) AND "Mem_Fer_FlancoCompleta" AND NOT "Mem_Fer_FlancoCompleta";   // rising edge of "Mem_Fer_FlancoCompleta"
   "Mem_Fer_FlancoCompleta" := "Mem_Fer_FlancoCompleta";
   IF #_w1 THEN "Alarmas".Fase_FermentacionTerminada := TRUE; END_IF;
END_REGION

REGION Network 5
   RUNG wire#powerrail
      Contact( "Alarmas".Fase_FermentacionTerminada )
      I_Contact( "ModoManual" )
      { S7_Templates := "SrcType := Real" } GT_Contact(in1 := "Fer_Volumen", in2 := "DatosDeRecetas".Fer_LimInfVolumen)
      S_Coil( "Act_BombaWash" )
   END_RUNG
   // the same network as SCL:
   IF "Alarmas".Fase_FermentacionTerminada AND NOT "ModoManual" AND ("Fer_Volumen" > "DatosDeRecetas".Fer_LimInfVolumen) THEN
       "Act_BombaWash" := TRUE;
   END_IF;
END_REGION

REGION Network 6
   RUNG wire#powerrail
      Contact( "Alarmas".Fase_FermentacionTerminada )
      { S7_Templates := "SrcType := Real" } LE_Contact(in1 := "Fer_Volumen", in2 := "DatosDeRecetas".Fer_LimInfVolumen)
      wire#w1
      R_Coil( "Alarmas".Fase_FermentacionTerminada )
   END_RUNG
   RUNG wire#w1
      S_Coil( "Alarmas".Fase_InicioLimpiezaFermentador )
   END_RUNG
   RUNG wire#w1
      S_Coil( "Alarmas".Fase_InicioDestilado )
   END_RUNG
   RUNG wire#w1
      R_Coil( "Alarmas".Fase_MomentoDescarteMetanol )
   END_RUNG
   // the same network as SCL:
   #_w1 := "Alarmas".Fase_FermentacionTerminada AND ("Fer_Volumen" <= "DatosDeRecetas".Fer_LimInfVolumen);
   IF #_w1 THEN
       "Alarmas".Fase_FermentacionTerminada := FALSE;
       "Alarmas".Fase_InicioLimpiezaFermentador := TRUE;
       "Alarmas".Fase_InicioDestilado := TRUE;
       "Alarmas".Fase_MomentoDescarteMetanol := FALSE;
   END_IF;
END_REGION

REGION Network 7
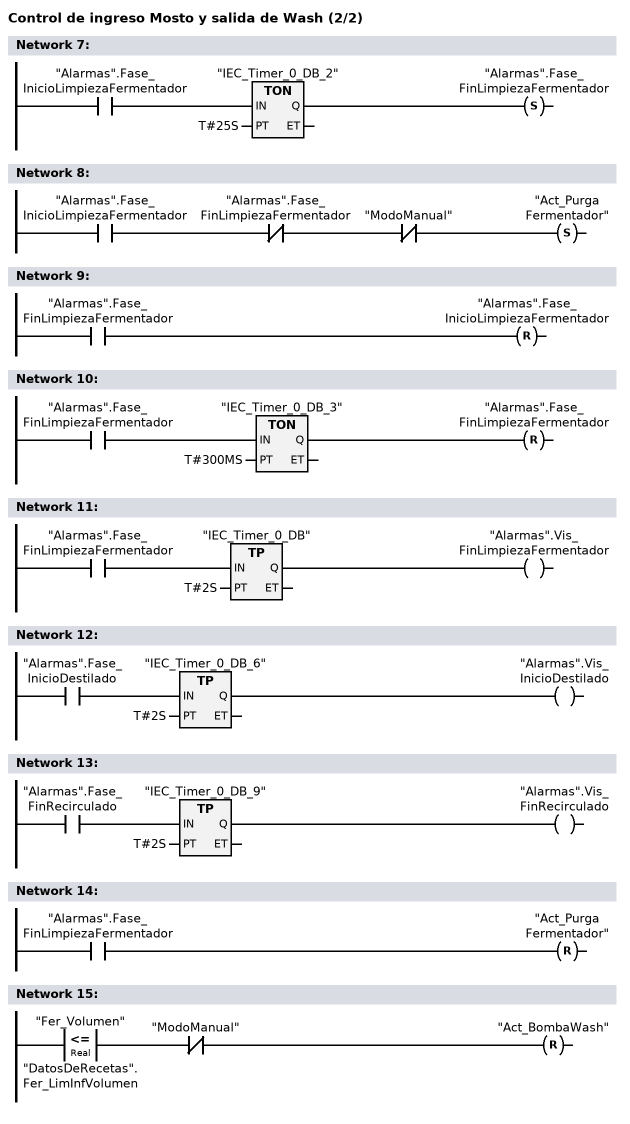
   "IEC_Timer_0_DB_2".TON(IN := "Alarmas".Fase_InicioLimpiezaFermentador, PT := T#25S);
   IF "IEC_Timer_0_DB_2".Q THEN "Alarmas".Fase_FinLimpiezaFermentador := TRUE; END_IF;
END_REGION

REGION Network 8
   RUNG wire#powerrail
      Contact( "Alarmas".Fase_InicioLimpiezaFermentador )
      I_Contact( "Alarmas".Fase_FinLimpiezaFermentador )
      I_Contact( "ModoManual" )
      S_Coil( "Act_PurgaFermentador" )
   END_RUNG
   // the same network as SCL:
   IF "Alarmas".Fase_InicioLimpiezaFermentador AND NOT "Alarmas".Fase_FinLimpiezaFermentador AND NOT "ModoManual" THEN
       "Act_PurgaFermentador" := TRUE;
   END_IF;
END_REGION

REGION Network 9
   RUNG wire#powerrail
      Contact( "Alarmas".Fase_FinLimpiezaFermentador )
      R_Coil( "Alarmas".Fase_InicioLimpiezaFermentador )
   END_RUNG
   // the same network as SCL:
   IF "Alarmas".Fase_FinLimpiezaFermentador THEN "Alarmas".Fase_InicioLimpiezaFermentador := FALSE; END_IF;
END_REGION

REGION Network 10
   "IEC_Timer_0_DB_3".TON(IN := "Alarmas".Fase_FinLimpiezaFermentador, PT := T#300MS);
   IF "IEC_Timer_0_DB_3".Q THEN "Alarmas".Fase_FinLimpiezaFermentador := FALSE; END_IF;
END_REGION

REGION Network 11
   "IEC_Timer_0_DB".TP(IN := "Alarmas".Fase_FinLimpiezaFermentador, PT := T#2S);
   "Alarmas".Vis_FinLimpiezaFermentador := "IEC_Timer_0_DB".Q;
END_REGION

REGION Network 12
   "IEC_Timer_0_DB_6".TP(IN := "Alarmas".Fase_InicioDestilado, PT := T#2S);
   "Alarmas".Vis_InicioDestilado := "IEC_Timer_0_DB_6".Q;
END_REGION

REGION Network 13
   "IEC_Timer_0_DB_9".TP(IN := "Alarmas".Fase_FinRecirculado, PT := T#2S);
   "Alarmas".Vis_FinRecirculado := "IEC_Timer_0_DB_9".Q;
END_REGION

REGION Network 14
   RUNG wire#powerrail
      Contact( "Alarmas".Fase_FinLimpiezaFermentador )
      R_Coil( "Act_PurgaFermentador" )
   END_RUNG
   // the same network as SCL:
   IF "Alarmas".Fase_FinLimpiezaFermentador THEN "Act_PurgaFermentador" := FALSE; END_IF;
END_REGION

REGION Network 15
   RUNG wire#powerrail
      { S7_Templates := "SrcType := Real" } LE_Contact(in1 := "Fer_Volumen", in2 := "DatosDeRecetas".Fer_LimInfVolumen)
      I_Contact( "ModoManual" )
      R_Coil( "Act_BombaWash" )
   END_RUNG
   // the same network as SCL:
   IF ("Fer_Volumen" <= "DatosDeRecetas".Fer_LimInfVolumen) AND NOT "ModoManual" THEN
       "Act_BombaWash" := FALSE;
   END_IF;
END_REGION
END_ORGANIZATION_BLOCK

ORGANIZATION_BLOCK "Control De Temperatura Del Fermentador"   // OB123, LAD, ProgramCycle
TITLE = "Main Program Sweep (Cycle)" / Control e la temperatura del Fermentador
{ S7_Optimized_Access := 'TRUE' }
VERSION : 0.1
// Nuestro fermentador solo tiene banda negativa; no tiene resistencia calefactora, solo refrigeración, esto tiene una razon de ser, al tratarse de una planta  en una zona cálida no se corre riesgo de que las levaduras mueran por el frío, si de calor y se avinagre el wash
   VAR_TEMP
      LimiteInferiorTemperatura : Real;
      LimiteSuperiorTemperatura : Real;
   END_VAR
   VAR_TEMP   // added for the SCL form of the ladder/FBD networks
      _w1 : Bool;
   END_VAR
BEGIN

REGION Network 1
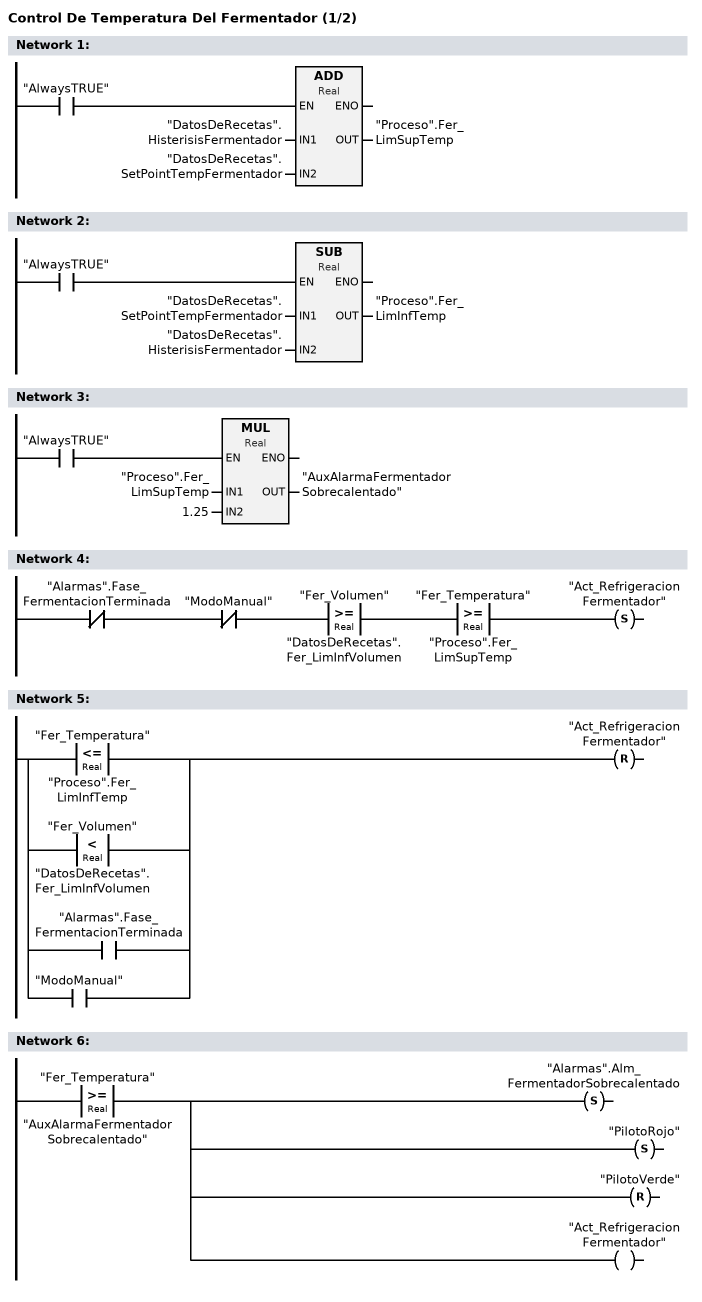
   RUNG wire#powerrail
      Contact( "AlwaysTRUE" )
      { S7_Templates := "SrcType := Real"; S7_GenerateENO := "TRUE" } Add(in1 := "DatosDeRecetas".HisterisisFermentador, in2 := "DatosDeRecetas".SetPointTempFermentador, out => "Proceso".Fer_LimSupTemp)
   END_RUNG
   // the same network as SCL:
   IF "AlwaysTRUE" THEN
       "Proceso".Fer_LimSupTemp := "DatosDeRecetas".HisterisisFermentador + "DatosDeRecetas".SetPointTempFermentador;
   END_IF;
END_REGION

REGION Network 2
   RUNG wire#powerrail
      Contact( "AlwaysTRUE" )
      { S7_Templates := "SrcType := Real"; S7_GenerateENO := "TRUE" } Sub(in1 := "DatosDeRecetas".SetPointTempFermentador, in2 := "DatosDeRecetas".HisterisisFermentador, out => "Proceso".Fer_LimInfTemp)
   END_RUNG
   // the same network as SCL:
   IF "AlwaysTRUE" THEN
       "Proceso".Fer_LimInfTemp := "DatosDeRecetas".SetPointTempFermentador - "DatosDeRecetas".HisterisisFermentador;
   END_IF;
END_REGION

REGION Network 3
   RUNG wire#powerrail
      Contact( "AlwaysTRUE" )
      { S7_Templates := "SrcType := Real"; S7_GenerateENO := "TRUE" } Mul(in1 := "Proceso".Fer_LimSupTemp, in2 := 1.25, out => "AuxAlarmaFermentadorSobrecalentado")
   END_RUNG
   // the same network as SCL:
   IF "AlwaysTRUE" THEN "AuxAlarmaFermentadorSobrecalentado" := "Proceso".Fer_LimSupTemp * 1.25; END_IF;
END_REGION

REGION Network 4
   RUNG wire#powerrail
      I_Contact( "Alarmas".Fase_FermentacionTerminada )
      I_Contact( "ModoManual" )
      { S7_Templates := "SrcType := Real" } GE_Contact(in1 := "Fer_Volumen", in2 := "DatosDeRecetas".Fer_LimInfVolumen)
      { S7_Templates := "SrcType := Real" } GE_Contact(in1 := "Fer_Temperatura", in2 := "Proceso".Fer_LimSupTemp)
      S_Coil( "Act_RefrigeracionFermentador" )
   END_RUNG
   // the same network as SCL:
   IF NOT "Alarmas".Fase_FermentacionTerminada AND NOT "ModoManual" AND ("Fer_Volumen" >= "DatosDeRecetas".Fer_LimInfVolumen) AND ("Fer_Temperatura" >= "Proceso".Fer_LimSupTemp) THEN
       "Act_RefrigeracionFermentador" := TRUE;
   END_IF;
END_REGION

REGION Network 5
   RUNG wire#powerrail
      { S7_Templates := "SrcType := Real" } LE_Contact(in1 := "Fer_Temperatura", in2 := "Proceso".Fer_LimInfTemp)
      wire#w1
      R_Coil( "Act_RefrigeracionFermentador" )
   END_RUNG
   RUNG wire#powerrail
      { S7_Templates := "SrcType := Real" } LT_Contact(in1 := "Fer_Volumen", in2 := "DatosDeRecetas".Fer_LimInfVolumen)
   END_RUNG wire#w1
   RUNG wire#powerrail
      Contact( "Alarmas".Fase_FermentacionTerminada )
   END_RUNG wire#w1
   RUNG wire#powerrail
      Contact( "ModoManual" )
   END_RUNG wire#w1
   // the same network as SCL:
   IF ("Fer_Temperatura" <= "Proceso".Fer_LimInfTemp) OR ("Fer_Volumen" < "DatosDeRecetas".Fer_LimInfVolumen) OR "Alarmas".Fase_FermentacionTerminada OR "ModoManual" THEN
       "Act_RefrigeracionFermentador" := FALSE;
   END_IF;
END_REGION

REGION Network 6
   RUNG wire#powerrail
      { S7_Templates := "SrcType := Real" } GE_Contact(in1 := "Fer_Temperatura", in2 := "AuxAlarmaFermentadorSobrecalentado")
      wire#w1
      S_Coil( "Alarmas".Alm_FermentadorSobrecalentado )
   END_RUNG
   RUNG wire#w1
      S_Coil( "PilotoRojo" )
   END_RUNG
   RUNG wire#w1
      R_Coil( "PilotoVerde" )
   END_RUNG
   RUNG wire#w1
      Coil( "Act_RefrigeracionFermentador" )
   END_RUNG
   // the same network as SCL:
   #_w1 := "Fer_Temperatura" >= "AuxAlarmaFermentadorSobrecalentado";
   IF #_w1 THEN
       "Alarmas".Alm_FermentadorSobrecalentado := TRUE;
       "PilotoRojo" := TRUE;
       "PilotoVerde" := FALSE;
   END_IF;
   "Act_RefrigeracionFermentador" := #_w1;
END_REGION

REGION Network 7
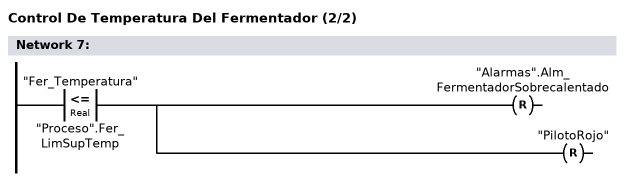
   RUNG wire#powerrail
      { S7_Templates := "SrcType := Real" } LE_Contact(in1 := "Fer_Temperatura", in2 := "Proceso".Fer_LimSupTemp)
      wire#w1
      R_Coil( "Alarmas".Alm_FermentadorSobrecalentado )
   END_RUNG
   RUNG wire#w1
      R_Coil( "PilotoRojo" )
   END_RUNG
   // the same network as SCL:
   IF "Fer_Temperatura" <= "Proceso".Fer_LimSupTemp THEN
       "Alarmas".Alm_FermentadorSobrecalentado := FALSE;
       "PilotoRojo" := FALSE;
   END_IF;
END_REGION
END_ORGANIZATION_BLOCK

// folder: Tanques

ORGANIZATION_BLOCK "Recirculado"   // OB125, LAD, ProgramCycle
TITLE = "Main Program Sweep (Cycle)"
{ S7_Optimized_Access := 'TRUE' }
VERSION : 0.1
   VAR_TEMP
      Impulso : Bool;
      InicioImpulso : Bool;
      Auxiliar : Real;
   END_VAR
   VAR CONSTANT
      Uno : Int := 1;
   END_VAR
   VAR_TEMP   // added for the SCL form of the ladder/FBD networks
      _w1 : Bool;
   END_VAR
BEGIN

REGION Network 1
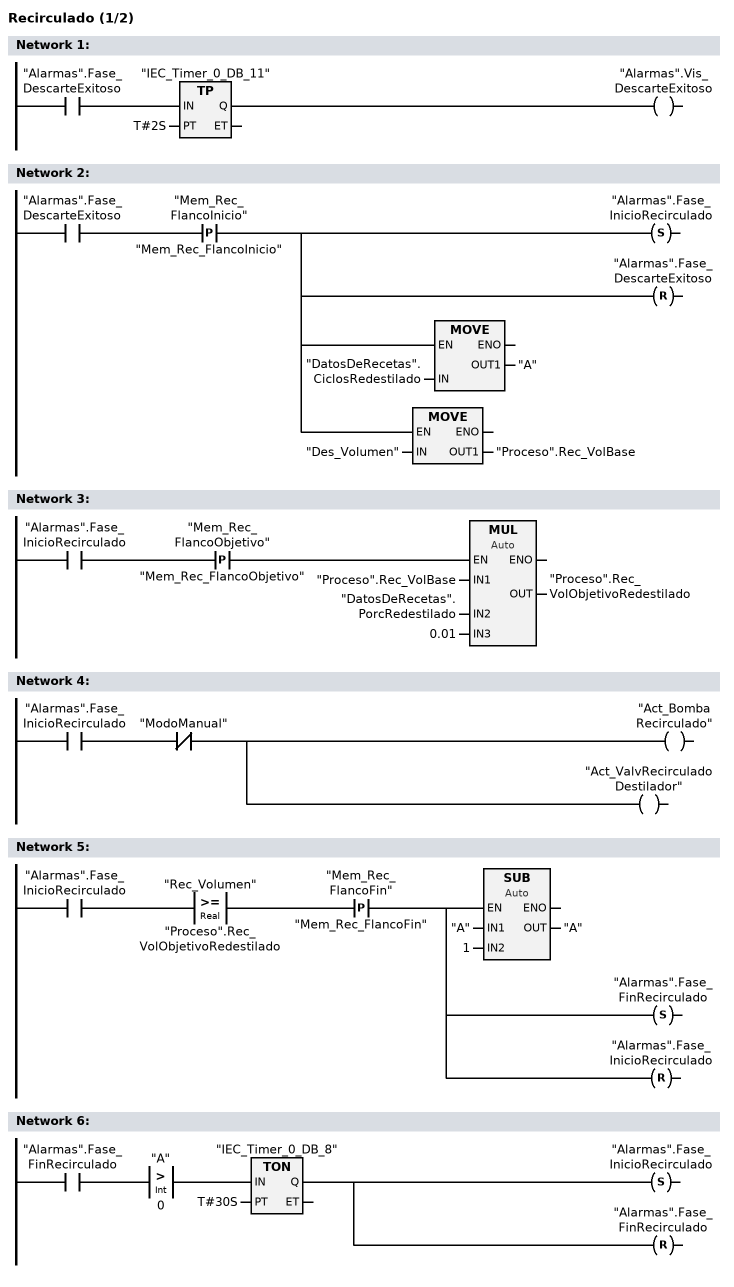
   "IEC_Timer_0_DB_11".TP(IN := "Alarmas".Fase_DescarteExitoso, PT := T#2S);
   "Alarmas".Vis_DescarteExitoso := "IEC_Timer_0_DB_11".Q;
END_REGION

REGION Network 2
   RUNG wire#powerrail
      Contact( "Alarmas".Fase_DescarteExitoso )
      P_Contact(operand := "Mem_Rec_FlancoInicio", bit := "Mem_Rec_FlancoInicio")
      wire#w1
      S_Coil( "Alarmas".Fase_InicioRecirculado )
   END_RUNG
   RUNG wire#w1
      R_Coil( "Alarmas".Fase_DescarteExitoso )
   END_RUNG
   RUNG wire#w1
      { S7_GenerateENO := "TRUE" } Move(in := "DatosDeRecetas".CiclosRedestilado, out1 => "A")
   END_RUNG
   RUNG wire#w1
      { S7_GenerateENO := "TRUE" } Move(in := "Des_Volumen", out1 => "Proceso".Rec_VolBase)
   END_RUNG
   // the same network as SCL:
   #_w1 := "Alarmas".Fase_DescarteExitoso AND "Mem_Rec_FlancoInicio" AND NOT "Mem_Rec_FlancoInicio";   // rising edge of "Mem_Rec_FlancoInicio"
   "Mem_Rec_FlancoInicio" := "Mem_Rec_FlancoInicio";
   IF #_w1 THEN
       "Alarmas".Fase_InicioRecirculado := TRUE;
       "Alarmas".Fase_DescarteExitoso := FALSE;
       "A" := "DatosDeRecetas".CiclosRedestilado;
       "Proceso".Rec_VolBase := "Des_Volumen";
   END_IF;
END_REGION

REGION Network 3
   RUNG wire#powerrail
      Contact( "Alarmas".Fase_InicioRecirculado )
      P_Contact(operand := "Mem_Rec_FlancoObjetivo", bit := "Mem_Rec_FlancoObjetivo")
      { S7_GenerateENO := "TRUE" } Mul(in1 := "Proceso".Rec_VolBase, in2 := "DatosDeRecetas".PorcRedestilado, in3 := 0.01, out => "Proceso".Rec_VolObjetivoRedestilado)
   END_RUNG
   // the same network as SCL:
   #_w1 := "Alarmas".Fase_InicioRecirculado AND "Mem_Rec_FlancoObjetivo" AND NOT "Mem_Rec_FlancoObjetivo";   // rising edge of "Mem_Rec_FlancoObjetivo"
   "Mem_Rec_FlancoObjetivo" := "Mem_Rec_FlancoObjetivo";
   IF #_w1 THEN
       "Proceso".Rec_VolObjetivoRedestilado := "Proceso".Rec_VolBase * "DatosDeRecetas".PorcRedestilado * 0.01;
   END_IF;
END_REGION

REGION Network 4
   RUNG wire#powerrail
      Contact( "Alarmas".Fase_InicioRecirculado )
      I_Contact( "ModoManual" )
      wire#w1
      Coil( "Act_BombaRecirculado" )
   END_RUNG
   RUNG wire#w1
      Coil( "Act_ValvRecirculadoDestilador" )
   END_RUNG
   // the same network as SCL:
   "Act_BombaRecirculado" := "Alarmas".Fase_InicioRecirculado AND NOT "ModoManual";
   "Act_ValvRecirculadoDestilador" := "Act_BombaRecirculado";
END_REGION

REGION Network 5
   RUNG wire#powerrail
      Contact( "Alarmas".Fase_InicioRecirculado )
      { S7_Templates := "SrcType := Real" } GE_Contact(in1 := "Rec_Volumen", in2 := "Proceso".Rec_VolObjetivoRedestilado)
      P_Contact(operand := "Mem_Rec_FlancoFin", bit := "Mem_Rec_FlancoFin")
      wire#w1
      { S7_GenerateENO := "TRUE" } Sub(in1 := "A", in2 := 1, out => "A")
   END_RUNG
   RUNG wire#w1
      S_Coil( "Alarmas".Fase_FinRecirculado )
   END_RUNG
   RUNG wire#w1
      R_Coil( "Alarmas".Fase_InicioRecirculado )
   END_RUNG
   // the same network as SCL:
   #_w1 := "Alarmas".Fase_InicioRecirculado AND ("Rec_Volumen" >= "Proceso".Rec_VolObjetivoRedestilado) AND "Mem_Rec_FlancoFin" AND NOT "Mem_Rec_FlancoFin";   // rising edge of "Mem_Rec_FlancoFin"
   "Mem_Rec_FlancoFin" := "Mem_Rec_FlancoFin";
   IF #_w1 THEN
       "A" := "A" - 1;
       "Alarmas".Fase_FinRecirculado := TRUE;
       "Alarmas".Fase_InicioRecirculado := FALSE;
   END_IF;
END_REGION

REGION Network 6
   "IEC_Timer_0_DB_8".TON(IN := "Alarmas".Fase_FinRecirculado AND ("A" > 0), PT := T#30S);
   IF "IEC_Timer_0_DB_8".Q THEN
       "Alarmas".Fase_InicioRecirculado := TRUE;
       "Alarmas".Fase_FinRecirculado := FALSE;
   END_IF;
END_REGION

REGION Network 7
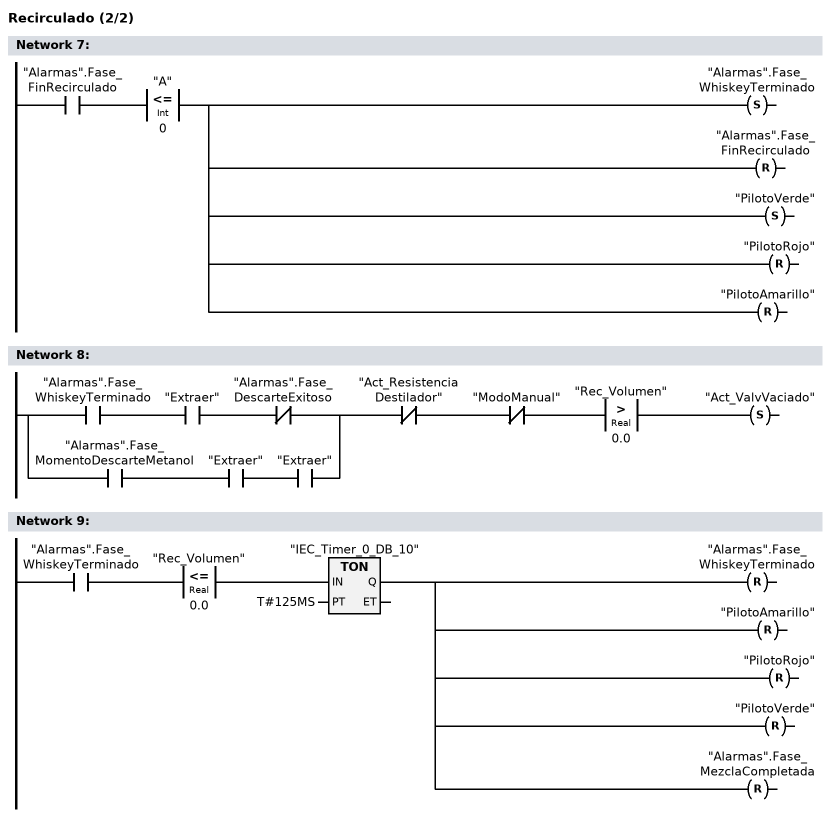
   RUNG wire#powerrail
      Contact( "Alarmas".Fase_FinRecirculado )
      { S7_Templates := "SrcType := Int" } LE_Contact(in1 := "A", in2 := 0)
      wire#w1
      S_Coil( "Alarmas".Fase_WhiskeyTerminado )
   END_RUNG
   RUNG wire#w1
      R_Coil( "Alarmas".Fase_FinRecirculado )
   END_RUNG
   RUNG wire#w1
      S_Coil( "PilotoVerde" )
   END_RUNG
   RUNG wire#w1
      R_Coil( "PilotoRojo" )
   END_RUNG
   RUNG wire#w1
      R_Coil( "PilotoAmarillo" )
   END_RUNG
   // the same network as SCL:
   IF "Alarmas".Fase_FinRecirculado AND ("A" <= 0) THEN "Alarmas".Fase_WhiskeyTerminado := TRUE; END_IF;
   #_w1 := "Alarmas".Fase_FinRecirculado AND ("A" <= 0);
   IF #_w1 THEN
       "Alarmas".Fase_FinRecirculado := FALSE;
       "PilotoVerde" := TRUE;
       "PilotoRojo" := FALSE;
       "PilotoAmarillo" := FALSE;
   END_IF;
END_REGION

REGION Network 8
   RUNG wire#powerrail
      Contact( "Alarmas".Fase_WhiskeyTerminado )
      Contact( "Extraer" )
      I_Contact( "Alarmas".Fase_DescarteExitoso )
      wire#w1
      I_Contact( "Act_ResistenciaDestilador" )
      I_Contact( "ModoManual" )
      { S7_Templates := "SrcType := Real" } GT_Contact(in1 := "Rec_Volumen", in2 := 0.0)
      S_Coil( "Act_ValvVaciado" )
   END_RUNG
   RUNG wire#powerrail
      Contact( "Alarmas".Fase_MomentoDescarteMetanol )
      Contact( "Extraer" )
      Contact( "Extraer" )
   END_RUNG wire#w1
   // the same network as SCL:
   IF (("Alarmas".Fase_WhiskeyTerminado AND "Extraer" AND NOT "Alarmas".Fase_DescarteExitoso) OR ("Alarmas".Fase_MomentoDescarteMetanol AND "Extraer" AND "Extraer")) AND NOT "Act_ResistenciaDestilador" AND NOT "ModoManual" AND ("Rec_Volumen" > 0.0) THEN
       "Act_ValvVaciado" := TRUE;
   END_IF;
END_REGION

REGION Network 9
   "IEC_Timer_0_DB_10".TON(IN := "Alarmas".Fase_WhiskeyTerminado AND ("Rec_Volumen" <= 0.0), PT := T#125MS);
   IF "IEC_Timer_0_DB_10".Q THEN
       "Alarmas".Fase_WhiskeyTerminado := FALSE;
       "PilotoAmarillo" := FALSE;
       "PilotoRojo" := FALSE;
       "PilotoVerde" := FALSE;
       "Alarmas".Fase_MezclaCompletada := FALSE;
   END_IF;
END_REGION
END_ORGANIZATION_BLOCK

(* ===== HMI "HMI_RT_1" =====
system functions are stored by id; their names below are inferred from use
connection "HMI_Conexión_1": ETHERNET, SMART_S7_1200_OMS

HMI tags "Variables del proceso"
   "DatosDeRecetas_SetPointTemperaturaAlambique" : Real = PLC DatosDeRecetas.SetPointTempDestilador AT %DB4.DBD266, 1 s
   "DatosDeRecetas_SetPointTemperaturaFermentador" : Real = PLC DatosDeRecetas.SetPointTempFermentador AT %DB4.DBD258, 1 s
   "DatosDeRecetas_HisterisisAlambique" : Real = PLC DatosDeRecetas.HisterisisDestilador AT %DB4.DBD270, 1 s
   "DatosDeRecetas_HisterisisFermentador" : Real = PLC DatosDeRecetas.HisterisisFermentador AT %DB4.DBD262, 1 s
   "DatosDeRecetas_PorcentajeDeAguaAgregada" : Real = PLC DatosDeRecetas.PorcAguaAgregada AT %DB4.DBD274, 1 s
   "DatosDeRecetas_PorcentajeDeVolumenEnPerdida" : Real = PLC DatosDeRecetas.PorcPerdidaDescarte AT %DB4.DBD282, 1 s
   "DatosDeRecetas_CiclosDeRefermentado" : Int = PLC DatosDeRecetas.CiclosRedestilado AT %DB4.DBW298, 1 s
   "DatosDeRecetas_PorcentaDeRedestilado" : Real = PLC DatosDeRecetas.PorcRedestilado AT %DB4.DBD278, 1 s
   "DatosDeRecetas_PorcentajePurgaFermentador" : Real = PLC DatosDeRecetas.PorcPurgaFermentador AT %DB4.DBD290, 1 s
   "DatosDeRecetas_PorcentajePurgaDestilador" : Real = PLC DatosDeRecetas.PorcPurgaDestilador AT %DB4.DBD294, 1 s
   "DatosDeRecetas_NombreReceta" : String[254] = PLC DatosDeRecetas.NombreReceta AT %DB4.DBX0.0, 1 s
   "DatosDeRecetas_NombreRecetaActiva" : Int = PLC DatosDeRecetas.NombreReceta_1 AT %DB4.DBW256, 1 s
   "DatosDeRecetas_VolumenDePerdida" : Real = PLC DatosDeRecetas.PorcPerdidaFermentacion AT %DB4.DBD286, 1 s
   "1- DB_Alarmas_FermentadorSobreCalentado" : Bool = PLC Alarmas.Alm_FermentadorSobrecalentado AT %DB6.DBX0.1, 1 s
   "ControlManual_ManualBombaDeWash" : Bool = PLC ControlManual.ManualBombaDeWash AT %DB2.DBX0.0, 1 s
   "ControlManual_ManualValvulaRecirculadoDestilador" : Bool = PLC ControlManual.ManualValvulaRecirculadoDestilador AT %DB2.DBX0.3, 1 s
   "ControlManual_ManualBombaDeAguaDestilador" : Bool = PLC ControlManual.ManualBombaDeAguaDestilador AT %DB2.DBX0.1, 1 s
   "ControlManual_ManualPurgaDestilador" : Bool = PLC ControlManual.ManualPurgaDestilador AT %DB2.DBX0.2, 1 s
   "ControlManual_ManualValvulaIngresoDeMosto" : Bool = PLC ControlManual.ManualValvulaIngresoDeMosto AT %DB2.DBX0.4, 1 s
   "ControlManual_ManualPurgaFermentador" : Bool = PLC ControlManual.ManualPurgaFermentador AT %DB2.DBX0.5, 1 s
   "ControlManual_ManualValvulaDeVaciado" : Bool = PLC ControlManual.ManualValvulaDeVaciado AT %DB2.DBX0.7, 1 s
   "ControlManual_ManualBombaDeRecirculado" : Bool = PLC ControlManual.ManualBombaDeRecirculado AT %DB2.DBX1.0, 1 s
   "DatosDeRecetas_Des_NivelBajo" : Real = PLC DatosDeRecetas.Des_NivelBajo AT %DB4.DBD316, 1 s
   "DatosDeRecetas_Des_LimSupVolumen" : Real = PLC DatosDeRecetas.Des_LimSupVolumen AT %DB4.DBD312, 1 s

HMI tags "Alambique"
   "TemperaturaAlambique" : Real = PLC Des_Temperatura AT %MD134, 500 ms
   "SetPointAlambique" : Real = PLC DatosDeRecetas.SetPointTempDestilador AT %DB4.DBD266, 500 ms
   "EstadoCalefactorAlambique" : Bool = PLC Act_ResistenciaDestilador AT %M36.4, 500 ms
   "PesoAlambique" : Real = PLC Des_Volumen AT %MD14, 500 ms
   "HisterisisTemperaturaAlambique" : Real = PLC DatosDeRecetas.HisterisisDestilador AT %DB4.DBD270, 500 ms
   "EstadoValvulaPurgaAlambique" : Bool = PLC Act_PurgaDestilador AT %M36.2, 500 ms
   "EstadoValvulaAguaAlambique" : Bool = PLC Act_BombaAguaDestilador AT %M36.1, 500 ms
   "EstadoBombaFermentadorAAlambique" : Bool = PLC Act_BombaWash AT %M36.0, 500 ms
   "EstadoBombaRecirculadoTanqueAAlambique" : Bool = PLC Act_ValvRecirculadoDestilador AT %M36.3, 500 ms
   "AlertaPesoAlambiqueBajo" : Bool = PLC AlertaAguaBajaDestilador AT %M132.3, 500 ms
   "NivelInferiorAlambique" : Bool = PLC NivelBajoDestiador AT %M132.4, 500 ms
   "LimiteSuperiorAlambique" : Bool = PLC Alarmas.Alm_DemasiadoWashDestilador AT %DB6.DBX0.4, 500 ms
   "FallaAlambique" : Bool = PLC AlertaAguaBajaDestilador AT %M132.3, 500 ms

HMI tags "Fermentador"
   "TemperaturaFermentador" : Real = PLC Fer_Temperatura AT %MD40, 500 ms
   "SetPointFermentador" : Real = PLC DatosDeRecetas.SetPointTempFermentador AT %DB4.DBD258, 500 ms
   "EstadoRefrigeracionFermentador" : Bool = PLC Act_RefrigeracionFermentador AT %M72.5, 500 ms
   "PesoFermentador" : Real = PLC Fer_Volumen AT %MD54, 500 ms
   "HisterisisTemperaturaFermentador" : Real = PLC DatosDeRecetas.HisterisisFermentador AT %DB4.DBD262, 500 ms
   "EstadoValvulaPurgaFermentador" : Bool = PLC Act_PurgaFermentador AT %M72.2, 500 ms
   "EstadoValvulaMosto" : Bool = PLC Act_ValvIngresoMosto AT %M72.1, 500 ms
   "NivelBajoFermentador" : Real = PLC DatosDeRecetas.Fer_LimInfVolumen AT %DB4.DBD304, 500 ms
   "NivelAltoFermentador" : Real = PLC DatosDeRecetas.Fer_LimSupVolumen AT %DB4.DBD308, 500 ms
   "FermentacionCompleta" : Bool = PLC Alarmas.Fase_FermentacionTerminada AT %DB6.DBX0.6, 500 ms
   "VolumenPerdida" : Real = PLC DatosDeRecetas.VolumenPerdida AT %DB4.DBD300, 500 ms

HMI tags "Tanques"
   "PesoTanqueRecirculado" : Real = PLC RecirVol AT %MD92, 500 ms
   "EstadoValvulaExtracccion" : Bool = PLC Act_ValvVaciado AT %M88.0, 500 ms
   "PesoTanqueRecepcion" : Real = PLC Rec_Volumen AT %MD82, 500 ms
   "EstadoValvulaRecirculado" : Bool = PLC Act_BombaRecirculado AT %M90.0, 500 ms

HMI tags "TablaNavegacion"
   "NumeroDeImagen" : Int, internal
   "NombreDeUsuario" : WString[10], internal
   "NombreImagen" : WString[10], internal

HMI tags "SistemaEnGeneral"
   "CiclosDeReDestilado" : Int, internal
   "PorcentajeDeAguaAñadida" : Real = PLC DatosDeRecetas.PorcAguaAgregada AT %DB4.DBD274, 1 s
   "ModoManualActivado" : Bool = PLC ModoManual AT %M500.0, 500 ms
   "ModoManualActivado_1" : Bool, internal
   "FermentacionTerminada" : Bool, internal
   "DestiladoTerminado" : Bool, internal
   "PorcentajeRedestilado" : Real = PLC DatosDeRecetas.PorcRedestilado AT %DB4.DBD278, 500 ms
   "NuevoSetPointAlambique" : Real, internal
   "IdDeReceta" : Int = PLC DatosDeRecetas.NombreReceta_1 AT %DB4.DBW256, 500 ms
   "AlarmasWord0" : Int AT %DB6.DBW0, 500 ms
   "AlarmasWord1" : Int AT %DB6.DBW1, 500 ms
   "Name" : String[254] = PLC DatosDeRecetas.NombreReceta AT %DB4.DBX0.0, 500 ms

HMI tags "Tabla de variables correccion"
   "AlarmasWord2" : Int AT %DB6.DBW4, 500 ms
   "NivelBajoDestilador" : Real AT %DB4.DBD316, 500 ms
   "LimSupDestilador" : Real AT %DB4.DBD312, 500 ms

discrete alarms
   2: 'Fermentador sobrecalentado: revisar refrigeracion', class Errors, trigger "AlarmasWord0" bit 9
   3: 'Aviso: Hay que descartar el metanol', class Errors, trigger "AlarmasWord0" bit 10
   4: 'Momento de descarte de metanol: presionar Extraer', class Errors, trigger "AlarmasWord0" bit 13
   5: 'Fermentador lleno: no puede ingresar más mosto', class Errors, trigger "AlarmasWord0" bit 11
   6: 'Fermentacion terminada', class Acknowledgement, trigger "AlarmasWord0" bit 14
   7: 'Inicio de limpieza del fermentador', class Acknowledgement, trigger "AlarmasWord0" bit 15
   8: 'Fin de limpieza del fermentador', class Acknowledgement, trigger "AlarmasWord2" bit 8
   9: 'Inicio de destilado', class Acknowledgement, trigger "AlarmasWord2" bit 9
   10: 'Inicio de clarificado', class Acknowledgement, trigger "AlarmasWord0" bit 2
   11: 'Demasiado wash en el destilador: purgar', class Warnings, trigger "AlarmasWord0" bit 12
   12: 'Descarte de metanol exitoso', class Acknowledgement, trigger "AlarmasWord2" bit 10
   13: 'Whiskey terminado: extraer producto', class Warnings, trigger "AlarmasWord0" bit 4
   14: 'Inicio de recirculado', class Acknowledgement, trigger "AlarmasWord0" bit 5
   15: 'Fin de recirculado', class Acknowledgement, trigger "AlarmasWord2" bit 11
   16: 'Mezcla completada', class Acknowledgement, trigger "AlarmasWord0" bit 7

analog alarms
   1: 'Destilador sin líquido: Calentamiento Apagado', class Errors, trigger "PesoAlambique"
   2: 'Demasiado Líquido en el alambique, favor de purgar para evitar cambios en la receta', class Warnings, trigger "PesoAlambique"
   3: 'El fermentador se encuentra lleno, no puede ingresar mas mosto y podría tardar mas de lo normal en refrigerarse', class Acknowledgement, trigger "PesoFermentador"
   4: 'El Fermentador tiene menos del nivel recomendable, refrigeración apagada', class Warnings, trigger "PesoFermentador"
   5: 'El Tanque de Recepción esta lleno, se frenará la destilación', class Errors, trigger "PesoTanqueRecepcion"
   6: 'El tanque de recirculado se llenó', class Acknowledgement, trigger "PesoTanqueRecirculadoPorcentual"

text list "Imagenes": 1 'Imagen raíz'; 2 'Home'; 4 'Imagen1'; 5 'Imagen2'; 6 'Imagen3'; 7 'Imágenes de sistema'; 8 'Diagnóstico de sistema SIMATIC PLC'; 9 'Tareas varias'; 10 'Administración de usuarios'; 11 'Información de sistema'; 12 'Tareas varias'; 13 ''; 14 ''; 15 ''; 16 ''; 17 'Imagen raíz'

recipe "Whiskey": NuevoSetPointAlambique <- "DatosDeRecetas_SetPointTemperaturaAlambique", NuevoSetPointFermentador <- "DatosDeRecetas_SetPointTemperaturaFermentador", NuevoHistAlambique <- "DatosDeRecetas_HisterisisAlambique", NuevoHistFermentador <- "DatosDeRecetas_HisterisisFermentador", NuevoPorcentajeAgua <- "DatosDeRecetas_PorcentajeDeAguaAgregada", NuevoVolumenPerdido <- "DatosDeRecetas_VolumenDePerdida", CiclosDeRedestilado <- "DatosDeRecetas_CiclosDeRefermentado", PorcentajeDeRedestilado <- "DatosDeRecetas_PorcentaDeRedestilado", PorcentajePurgaFermentador <- "DatosDeRecetas_PorcentajePurgaFermentador", PorcentajePurgaDestilador <- "DatosDeRecetas_PorcentajePurgaDestilador", NombreDeRegistro <- "DatosDeRecetas_NombreReceta", IdDeReceta <- "IdDeReceta"

screen "Home" 320x240, template "con fondo"
   on GenerateScreen: SetTag("NombreImagen", 'Home')
   TextField "Campo de texto_1" at 62,43 size 60x13; Text 'Bienvenido,'
   IOField "Campo ES_1" at 118,39 size 96x23; FormatPattern ????????????
      ProcessValue <- "NombreDeUsuario"
   Button "Botón_1" at 26,69 size 68x33; TextOff 'Vista General'; Authorization "Monitorización"
      on Release: ActivateScreen("Vista General", 0)
   Button "Botón_2" at 117,68 size 75x32; TextOff 'Fermentador'; Authorization "Monitorización"
      on Release: ActivateScreen("Fermentador", 0)
   Button "Botón_3" at 214,68 size 68x32; TextOff 'Destilador'; Authorization "Monitorización"
      on Release: ActivateScreen("Alambique", 0)
   Button "Botón_4" at 116,111 size 75x30; TextOff 'Explicación'
      on Release: ActivateScreen("explicacion", 0)
   Button "Botón_5" at 25,111 size 69x32; TextOff 'Tanques'; Authorization "Monitorización"
      on Release: ActivateScreen("Tanques", 0)
   Button "Botón_6" at 213,112 size 69x29; TextOff 'Configuración'; Authorization "Operación"
      on Release: ActivateScreen("Configuración", 0)
   Button "Botón_7" at 72,155 size 64x32; TextOff 'Estadísticas'; Authorization "Monitorización"
   Button "Botón_8" at 177,155 size 57x31; TextOff 'Alarmas'; Authorization "Monitorización"
      on Release: ActivateScreen("Alarmas", 0)

screen "Vista General" 320x240, template "con fondo"
   on GenerateScreen: SetTag("NombreImagen", 'Vista General')
   TextField "Campo de texto_1" at 169,187 size 62x15; Text 'Alambique'
   GraphicView "Visor de gráficos_2" at 196,30 size 81x143; Picture "torre_destilacion"
   TextField "Campo de texto_2" at 10,187 size 76x15; Text 'Fermentador'
   IOField "Campo ES_4" at 115,171 size 47x14; Authorization "Monitorización"; FormatPattern s999.99; Unit °C
      ProcessValue <- "TemperaturaFermentador"
   TextField "Campo de texto_11" at 93,189 size 19x15; Text 'SP:'
   IOField "Campo ES_2" at 115,191 size 47x14; Authorization "Monitorización"; FormatPattern s999.99; Unit °C
      ProcessValue <- "SetPointFermentador"
   IOField "Campo ES_3" at 270,172 size 49x14; Authorization "Monitorización"; FormatPattern s999.999; Unit °C
      ProcessValue <- "TemperaturaAlambique"
   TextField "Campo de texto_4" at 254,172 size 12x15; Text 'T:'
   TextField "Campo de texto_6" at 247,190 size 19x15; Text 'SP:'
   IOField "Campo ES_5" at 270,192 size 49x14; Authorization "Monitorización"; FormatPattern s999.999; Unit °C
      ProcessValue <- "SetPointAlambique"
   GraphicView "Visor de gráficos_3" at 185,139 size 36x30; Picture "valvula_abierta"
   GraphicView "Visor de gráficos_5" at 252,99 size 36x30; Picture "valvula_abierta"
   TextField "Campo de texto_3" at 189,162 size 32x13; Text 'Purga'
   TextField "Campo de texto_5" at 178,83 size 28x13; Text 'Wash'
   GraphicView "Visor de gráficos_6" at 185,95 size 36x30; Picture "valvula_abierta"
   GraphicView "Visor de gráficos_7" at 45,40 size 64x135; Picture "fermentador_con_serpentin"
   GraphicView "Visor de gráficos_9" at 18,53 size 36x30; Picture "valvula_abierta"
   TextField "Campo de texto_9" at 14,81 size 32x13; Text 'Mosto'
   GraphicView "Visor de gráficos_10" at 18,139 size 36x30; Picture "valvula_abierta"
   TextField "Campo de texto_12" at 22,169 size 32x13; Text 'Purga'
      Visibility <- "EstadoValvulaPurgaFermentador"
   GraphicView "Visor de gráficos_12" at 109,82 size 29x27; Picture "Gráfico_9"
      Visibility <- "EstadoRefrigeracionFermentador"
   GraphicView "Visor de gráficos_8" at 178,50 size 32x31; Picture "Gráfico_10"
   Line "Línea_1" at 223,149 size 0x10
      Appearance <- "EstadoCalefactorAlambique"
   Line "Línea_2" at 224,159 size 25x0
      Appearance <- "EstadoCalefactorAlambique"
   Line "Línea_3" at 223,149 size 3x6
      Appearance <- "EstadoCalefactorAlambique"
   Line "Línea_4" at 227,150 size 3x5
      Appearance <- "EstadoCalefactorAlambique"
   Line "Línea_5" at 230,150 size 3x5
      Appearance <- "EstadoCalefactorAlambique"
   Line "Línea_6" at 233,150 size 3x5
      Appearance <- "EstadoCalefactorAlambique"
   Line "Línea_7" at 236,150 size 3x5
      Appearance <- "EstadoCalefactorAlambique"
   Line "Línea_8" at 239,150 size 3x5
      Appearance <- "EstadoCalefactorAlambique"
   Line "Línea_9" at 242,150 size 3x5
      Appearance <- "EstadoCalefactorAlambique"
   Line "Línea_10" at 245,150 size 3x5
      Appearance <- "EstadoCalefactorAlambique"
   GraphicView "Visor de gráficos_13" at 178,49 size 34x33; Picture "Gráfico_12"
      Visibility <- "EstadoBombaFermentadorAAlambique"
   GraphicView "Visor de gráficos_14" at 253,100 size 36x31; Picture "valvula_cerrada"
      Visibility <- "EstadoBombaRecirculadoTanqueAAlambique"
   GraphicView "Visor de gráficos_4" at 103,48 size 78x33; Picture "Gráfico_11"
   TextField "Campo de texto_7" at 259,84 size 57x15; Text 'Recirculado'
   GraphicView "Visor de gráficos_15" at 185,95 size 36x31; Picture "valvula_cerrada"
      Visibility <- "EstadoValvulaAguaAlambique"
   TextField "Campo de texto_8" at 189,117 size 28x13; Text 'Agua'
   GraphicView "Visor de gráficos_16" at 185,135 size 36x31; Picture "valvula_cerrada"
      Visibility <- "EstadoValvulaPurgaAlambique"
   GraphicView "Visor de gráficos_17" at 14,139 size 36x31; Picture "valvula_cerrada"
      Visibility <- "EstadoValvulaPurgaFermentador"
   GraphicView "Visor de gráficos_18" at 18,53 size 36x31; Picture "valvula_cerrada"
      Visibility <- "EstadoValvulaMosto"
   TextField "Campo de texto_10" at 100,170 size 12x15; Text 'T:'
   Button "Botón_3" at 14,50 size 36x31; TextOff 'Text'
      on Release: InvertBit("ControlManual_ManualValvulaIngresoDeMosto")
   Button "Botón_2" at 12,138 size 38x32; TextOff 'Text'
      on Release: InvertBit("ControlManual_ManualPurgaFermentador")
   Button "Botón_6" at 170,40 size 47x45; TextOff 'Text'
      on Press: InvertBit("ControlManual_ManualBombaDeWash")
   Button "Botón_1" at 184,94 size 38x32; TextOff 'Text'
      on Release: InvertBit("ControlManual_ManualBombaDeAguaDestilador")
   Button "Botón_4" at 177,135 size 45x27; TextOff 'Text'
      on Release: InvertBit("ControlManual_ManualPurgaDestilador")
   Button "Botón_5" at 254,98 size 39x28; TextOff 'Text'
      on Press: InvertBit("ControlManual_ManualValvulaRecirculadoDestilador")

screen "P&id" 320x240, template "con fondo"
   on GenerateScreen: SetTag("NombreImagen", 'Diagrama P&ID')
   GraphicView "Visor de gráficos_1" at 10,51 size 305x155; Picture "pid_completo"

screen "Alarmas" 320x240, template "con fondo"
   on GenerateScreen: SetTag("NombreImagen", 'Alarma')
   AlarmView "Visor de avisos_1" at 18,33 size 261x168

screen "Información del proyecto" 320x240, template "con fondo"
   on GenerateScreen: SetTag("NombreImagen", 'Información')
   TextField "HmiScreenItemData" at 57,71 size 98x20; Text 'Nombre del proyecto:'
   TextField "HmiScreenItemData_1" at 159,71 size 157x20; Text 'Conjunto destiladora-fermentador'
   TextField "HmiScreenItemData_2" at 57,92 size 98x20; Text 'Creado:'
   TextField "HmiScreenItemData_3" at 159,92 size 157x20; Text '04/10/2026 1:18:15'
   TextField "HmiScreenItemData_4" at 57,113 size 98x20; Text 'Autor:'
   TextField "HmiScreenItemData_5" at 159,113 size 157x20; Text 'nalbert'
   TextField "HmiScreenItemData_6" at 57,134 size 98x20; Text 'Descripción:'
   TextField "HmiScreenItemData_7" at 159,134 size 157x20; Text '(no configurado)'

screen "Administración de usuarios" 320x240, template "con fondo"
   on GenerateScreen: SetTag("NombreImagen", 'Control de Usuarios')
   UserView "HmiScreenItemData" at 57,39 size 263x163

screen "Información de sistema" 320x240, template "con fondo"
   on GenerateScreen: SetTag("NombreImagen", 'Información')
   TextField "HmiScreenItemData" at 57,71 size 98x20; Text 'Tipo de panel:'
   TextField "HmiScreenItemData_1" at 159,71 size 157x20; Text 'KTP600 Basic color PN 12.0'
   TextField "HmiScreenItemData_2" at 57,92 size 98x20; Text 'Conexión:'
   TextField "HmiScreenItemData_3" at 159,92 size 157x20; Text '(no configurado)'
   TextField "HmiScreenItemData_4" at 57,113 size 98x20; Text 'Controlador:'
   TextField "HmiScreenItemData_5" at 159,113 size 157x20; Text '<PLC>'

Template "con fondo" 320x240
   Button "Imagen inicial" at 14,211 size 35x29; TextOff 'Imagen inicial'; PictureOff "NavigateHome_KTP600_Basic_color_PN"; PictureOn "NavigateHome_KTP600_Basic_color_PN"
      on Release: ActivateScreen("Home", 0)
   Button "Iniciar sesión" at 222,211 size 36x29; TextOff 'Iniciar sesión'; PictureOff "Login_KTP600_Basic_color_PN"; PictureOn "Login_KTP600_Basic_color_PN"; Authorization "Administración de usuarios"
      on Release: ActivateScreen("Administración de usuarios", 0)
   Button "Idioma" at 116,210 size 38x29; TextOff 'Idioma'; PictureOn "ToggleLanguage_KTP600_Basic_color_PN"; PictureOff "boton_graficos_64"
      on Release: ActivateScreen("estadisticas", 0)
   Button "Avisos" at 167,211 size 39x28; TextOff 'Avisos'; PictureOff "AlarmDisplay_KTP600_Basic_color_PN"; PictureOn "AlarmDisplay_KTP600_Basic_color_PN"
      on Release: ActivateScreen("Alarmas", 0)
   Button "Salir" at 270,210 size 38x29; TextOff 'Salir'; PictureOff "ExitRuntime_KTP600_Basic_color_PN"; PictureOn "ExitRuntime_KTP600_Basic_color_PN"; Authorization "Monitorización"
      on Release: function_f23ef4c9()
   DateTimeField "HmiScreenItemData" at 223,16 size 85x19
   DateTimeField "HmiScreenItemData_1" at 235,0 size 85x19
   GraphicView "Logotipo" at 0,0 size 106x38; Picture "Logotipo de HMI_1"
   Button "Plantilla_Botón_1" at 67,210 size 35x29; TextOff '?'; PictureOff "Left_Arrow"
      on Release: ActivateScreen("explicacion", 0)
   IOField "Plantilla_Campo ES_1" at 113,4 size 135x26; FormatPattern ??????????????????????
      ProcessValue <- "NombreImagen"
   Softkey "Softkey_F1" at 0,0 size 0x0
      on KeyUp: ActivateScreen("Home", 0)
   Softkey "Softkey_F2" at 0,0 size 0x0
      on KeyUp: ActivateScreen("explicacion", 0)
   Softkey "Softkey_F3" at 0,0 size 0x0
      on KeyUp: ActivateScreen("estadisticas", 0)
   Softkey "Softkey_F4" at 0,0 size 0x0
      on KeyUp: ActivateScreen("Alarmas", 0)
   Softkey "Softkey_F5" at 0,0 size 0x0
      on KeyUp: ActivateScreen("Administración de usuarios", 0)
   Softkey "Softkey_F6" at 0,0 size 0x0
      on KeyUp: ActivateScreen("inicio", 0)

screen "inicio" 320x240
   GraphicView "Visor de gráficos_1" at 78,14 size 151x99; Picture "etiqueta_whiskey_borde"
   TextField "Campo de texto_1" at 8,115 size 134x13; Text 'Proyecto Final de SCADA:'
   TextField "Campo de texto_2" at 94,126 size 226x13; Text 'Conjunto fermentador- destileria de Whiskey'
   TextField "Campo de texto_3" at 11,140 size 43x13; Text 'Alumno:'
   TextField "Campo de texto_4" at 94,139 size 101x13; Text 'Fabricio David Gallo'
   TextField "Campo de texto_5" at 11,158 size 60x13; Text 'Profesores:'
   TextField "Campo de texto_6" at 94,158 size 187x13; Text 'Ing Daniel Gamero, Lic.Julian Minatel'
   Button "Botón_1" at 59,189 size 192x42; TextOff 'Click aquí para iniciar'; Authorization "Monitorización"
      on Click: function_f41c6f6c("NombreDeUsuario"); ActivateScreen("Home", 0)

screen "Fermentador" 320x240, template "con fondo"
   on GenerateScreen: SetTag("NombreImagen", 'Fermentador')
   TextField "Campo de texto_2" at 115,39 size 67x13; Text 'Fermentador'
   IOField "Campo ES_4" at 257,69 size 48x14; Authorization "Monitorización"; FormatPattern s99.999; Unit °C
      ProcessValue <- "SetPointFermentador"
   TextField "Campo de texto_10" at 113,51 size 71x13; Text 'Temperatura:'
   TextField "Campo de texto_11" at 233,68 size 18x13; Text 'SP:'
   IOField "Campo ES_2" at 185,53 size 54x14; Authorization "Monitorización"; FormatPattern s999.999; Unit °C
      ProcessValue <- "TemperaturaFermentador"
   TextField "Campo de texto_5" at 123,150 size 28x13; Text 'Wash'
   GraphicView "Visor de gráficos_7" at 45,40 size 64x135; Picture "fermentador_con_serpentin"
   GraphicView "Visor de gráficos_9" at 18,53 size 36x30; Picture "valvula_abierta"
   TextField "Campo de texto_9" at 14,81 size 32x13; Text 'Mosto'
   GraphicView "Visor de gráficos_10" at 18,139 size 36x30; Picture "valvula_abierta"
   TextField "Campo de texto_12" at 22,169 size 32x13; Text 'Purga'
   GraphicView "Visor de gráficos_12" at 18,100 size 29x27; Picture "Gráfico_9"
      Visibility <- "EstadoRefrigeracionFermentador"
   GraphicView "Visor de gráficos_8" at 123,127 size 29x26; Picture "Gráfico_10"
   GraphicView "Visor de gráficos_13" at 124,127 size 31x26; Picture "Gráfico_12"
      Visibility <- "EstadoBombaFermentadorAAlambique"
   GraphicView "Visor de gráficos_17" at 14,139 size 36x31; Picture "valvula_cerrada"
      Visibility <- "ControlManual_ManualPurgaFermentador"
   GraphicView "Visor de gráficos_18" at 18,53 size 36x31; Picture "valvula_cerrada"
      Visibility <- "EstadoValvulaMosto"
   GraphicView "Visor de gráficos_1" at 102,125 size 22x32; Picture "Gráfico_24"
   TextField "Campo de texto_1" at 113,67 size 52x13; Text 'Histerisis:'
   TextField "Campo de texto_3" at 113,83 size 73x13; Text 'Nivel Inferior:'
   TextField "Campo de texto_4" at 114,95 size 75x13; Text 'Nivel superior:'
   TextField "Campo de texto_6" at 135,182 size 105x13; Text 'Volumen de Pérdida:'
   Button "Botón_1" at 277,36 size 38x24; TextOff 'Text'; PictureOff "Gráfico_13"
      on Release: ActivateScreen("Alambique", 0)
   IOField "Campo ES_1" at 184,70 size 42x14; Authorization "Monitorización"; FormatPattern s99.99; Unit °C
      ProcessValue <- "HisterisisTemperaturaFermentador"
   IOField "Campo ES_3" at 203,85 size 71x14; Authorization "Monitorización"; FormatPattern s999.999; Unit L
      ProcessValue <- "NivelBajoFermentador"
   IOField "Campo ES_5" at 203,99 size 71x14; Authorization "Monitorización"; FormatPattern s999.999; Unit L
      ProcessValue <- "NivelAltoFermentador"
   TextField "Campo de texto_7" at 155,122 size 66x15; Text 'Alambique'
   TextField "Campo de texto_8" at 148,163 size 83x13; Text 'Volumen Actual:'
   Button "Botón_2" at 12,137 size 38x32; TextOff 'Text'
      on Release: InvertBit("ControlManual_ManualPurgaFermentador")
   Button "Botón_3" at 10,49 size 40x34; TextOff 'Text'
      on Release: InvertBit("ControlManual_ManualValvulaIngresoDeMosto")
   Button "Botón_4" at 116,120 size 54x42; TextOff 'Text'
      on Release: InvertBit("ControlManual_ManualBombaDeWash")
   IOField "Campo ES_6" at 240,162 size 71x14; FormatPattern s999999999.999; Unit L
      ProcessValue <- "PesoFermentador"
   IOField "Campo ES_7" at 240,181 size 71x14; FormatPattern s99999; Unit %
      ProcessValue <- "VolumenPerdida"

screen "Alambique" 320x240, template "con fondo"
   on GenerateScreen: SetTag("NombreImagen", 'Destilador')
   GraphicView "Visor de gráficos_2" at 29,41 size 95x157; Picture "torre_destilacion"
   TextField "Campo de texto_1" at 10,38 size 55x13; Text 'Alambique'
   IOField "Campo ES_3" at 270,68 size 42x14; Authorization "Monitorización"; FormatPattern 999.9; Unit °C
   TextField "Campo de texto_4" at 203,66 size 68x13; Text 'Temperatura'
   TextField "Campo de texto_6" at 244,85 size 18x13; Text 'SP:'
   IOField "Campo ES_5" at 270,85 size 42x14; Authorization "Monitorización"; FormatPattern 999.9; Unit °C
   GraphicView "Visor de gráficos_3" at 96,154 size 36x33; Picture "valvula_abierta"
   TextField "Campo de texto_5" at 6,94 size 28x13; Text 'Wash'
   GraphicView "Visor de gráficos_6" at 6,160 size 37x34; Picture "valvula_abierta"
   GraphicView "Visor de gráficos_8" at 6,63 size 32x31; Picture "Gráfico_10"
   GraphicView "Visor de gráficos_13" at 6,63 size 34x31; Picture "Gráfico_12"
      Visibility <- "EstadoBombaFermentadorAAlambique"
   GraphicView "Visor de gráficos_15" at 96,154 size 36x31; Picture "valvula_cerrada"
      Visibility <- "EstadoValvulaPurgaAlambique"
   TextField "Campo de texto_8" at 10,188 size 28x13; Text 'Agua'
   GraphicView "Visor de gráficos_16" at 6,159 size 40x34; Picture "valvula_cerrada"
      Visibility <- "EstadoValvulaAguaAlambique"
   TextField "Campo de texto_2" at 119,53 size 72x15; Text '> Al tanque'
   TextField "Campo de texto_3" at 106,174 size 32x13; Text 'Purga'
   TextField "Campo de texto_9" at 136,82 size 76x15; Text '<Del tanque'
   GraphicView "Visor de gráficos_4" at 96,74 size 39x33; Picture "valvula_abierta"
   GraphicView "Visor de gráficos_14" at 96,76 size 40x30; Picture "valvula_cerrada"
      Visibility <- "EstadoValvulaRecirculado"
   Button "Botón_1" at 284,34 size 25x23; TextOff 'Text'; PictureOff "Gráfico_13"
      on Release: ActivateScreen("Tanques", 0)
   Button "Botón_5" at 252,34 size 26x23; TextOff 'Text'; PictureOff "Gráfico_14"
      on Release: function_efd93a16()
   TextField "Campo de texto_7" at 99,97 size 60x13; Text 'Recirculado'
   TextField "Campo de texto_10" at 180,119 size 83x13; Text 'Volumen Actual:'
   IOField "Campo ES_2" at 271,121 size 41x17; Authorization "Monitorización"; FormatPattern 999.9; Unit L
   TextField "Campo de texto_12" at 219,99 size 52x13; Text 'Histerisis:'
   TextField "Campo de texto_13" at 169,139 size 73x13; Text 'Nivel Inferior:'
   TextField "Campo de texto_14" at 169,157 size 75x13; Text 'Nivel superior:'
   IOField "Campo ES_1" at 271,102 size 42x14; Authorization "Monitorización"; FormatPattern 999.9; Unit °C
   IOField "Campo ES_6" at 247,140 size 42x14; Authorization "Monitorización"; FormatPattern 999.9; Unit L
   IOField "Campo ES_7" at 247,156 size 42x14; Authorization "Monitorización"; FormatPattern 999.9; Unit L
   Button "Botón_3" at 3,159 size 48x32; TextOff 'Text'
      on Release: InvertBit("ControlManual_ManualBombaDeAguaDestilador")
   Button "Botón_2" at 101,152 size 45x27; TextOff 'Text'
      on Release: InvertBit("ControlManual_ManualPurgaDestilador")
   Button "Botón_4" at 99,74 size 39x28; TextOff 'Text'
      on Press: InvertBit("ControlManual_ManualValvulaRecirculadoDestilador")
   Button "Botón_6" at 6,57 size 45x40; TextOff 'Text'
      on Press: InvertBit("ControlManual_ManualBombaDeWash")

screen "Tanques" 320x240, template "con fondo"
   on GenerateScreen: SetTag("NombreImagen", 'Tanques')
   GraphicView "Visor de gráficos_1" at 41,37 size 68x107; Picture "Gráfico_22"
   GraphicView "Visor de gráficos_8" at 150,160 size 40x34; Picture "Gráfico_10"
   GraphicView "Visor de gráficos_2" at 137,86 size 53x54; Picture "Gráfico_22"
   GraphicView "Visor de gráficos_4" at 0,47 size 47x33; Picture "Gráfico_24"
   GraphicView "Visor de gráficos_13" at 150,159 size 41x36; Picture "Gráfico_12"
      Visibility <- "EstadoBombaRecirculadoTanqueAAlambique"
   GraphicView "Visor de gráficos_5" at 104,97 size 36x30; Picture "valvula_abierta"
   GraphicView "Visor de gráficos_3" at 104,95 size 36x31; Picture "valvula_cerrada"
      Visibility <- "EstadoValvulaRecirculado"
   GraphicView "Visor de gráficos_6" at 150,136 size 32x25; Picture "Gráfico_25"
   GraphicView "Visor de gráficos_9" at 58,136 size 39x37; Picture "valvula_abierta_2"
   GraphicView "Visor de gráficos_10" at 58,136 size 38x40; Picture "valvula_cerrada_1"
      Visibility <- "EstadoValvulaExtracccion"
   TextField "Campo de texto_1" at 54,176 size 50x15; Text 'Vaciado'
   TextField "Campo de texto_2" at 191,156 size 66x15; Text 'Alambique'
   TextField "Campo de texto_3" at 110,37 size 60x15; Text 'Recepción'
   TextField "Campo de texto_4" at 196,80 size 68x15; Text 'Recirculado'
   TextField "Campo de texto_5" at 110,51 size 32x15; Text 'Peso:'
   TextField "Campo de texto_6" at 196,95 size 32x15; Text 'Peso:'
   Button "Botón_5" at 276,38 size 40x27; TextOff 'Text'; PictureOff "Gráfico_14"
      on Release: function_efd93a16()
   IOField "Campo ES_1" at 241,97 size 75x14; FormatPattern s999.999; Unit L
      ProcessValue <- "PesoTanqueRecirculado"
   IOField "Campo ES_2" at 150,53 size 75x14; FormatPattern s999.99; Unit L
      ProcessValue <- "PesoTanqueRecepcion"
   Button "Botón_2" at 109,97 size 31x26; TextOff 'Text'
      on Release: InvertBit("ControlManual_ManualValvulaRecirculadoDestilador")
   Button "Botón_1" at 51,129 size 58x55; TextOff 'Text'
      on Release: InvertBit("ControlManual_ManualValvulaDeVaciado")
   Button "Botón_3" at 146,152 size 63x46; TextOff 'Text'
      on Release: InvertBit("ControlManual_ManualBombaDeRecirculado")

screen "explicacion" 320x240, template "con fondo"
   on GenerateScreen: SetTag("NombreImagen", 'Detalle')
   TextField "Campo de texto_1" at 16,48 size 261x13; Text 'El sistema comprende tres etapas diferenciadas: Fermentador,'
   TextField "Campo de texto_2" at 25,62 size 251x13; Text 'destilador (/alambique) y el sistema de tanques y extracción.'
   Button "Botón_1" at 26,83 size 252x25; TextOff 'Puedes ver el diagrama P&ID del proceso completo aquí'
      on Release: ActivateScreen("P&id", 0)
   Button "Botón_2" at 26,113 size 252x25; TextOff 'Información detallada de cada etapa'
      on Release: ActivateScreen("Información de sistema", 0)
   Button "Botón_3" at 26,176 size 252x25; TextOff 'Como operar los botones inferiores'
      on Release: ActivateScreen("explicacion botones inferiores", 0)
   Button "Botón_4" at 26,143 size 252x25; TextOff 'Información del proyecto'
      on Release: ActivateScreen("Información del proyecto", 0)
   Button "Botón_5" at 278,48 size 40x27; TextOff 'Text'; PictureOff "Gráfico_14"
      on Release: ActivateScreen("Home", 0)

screen "explicacion botones inferiores" 320x240, template "con fondo"
   TextField "Campo de texto_1" at 12,46 size 89x12; Text 'Con este botón volvés'
   TextField "Campo de texto_2" at 12,58 size 84x12; Text 'a la pantalla de inicio'
   TextField "Campo de texto_3" at 162,42 size 95x12; Text 'Con este botón accedés'
   TextField "Campo de texto_4" at 160,54 size 101x12; Text 'al menú de explicaciones'
   TextField "Campo de texto_5" at 180,79 size 95x12; Text 'Con este botón accedés'
   TextField "Campo de texto_6" at 178,91 size 101x12; Text 'al menú de explicaciones'
   TextField "Campo de texto_7" at 153,112 size 121x12; Text 'Acá están las alarmas y avisos'
   TextField "Campo de texto_8" at 205,134 size 77x12; Text 'Control de usuarios'
   TextField "Campo de texto_9" at 265,155 size 45x12; Text 'Cerrar HMI'

screen "estadisticas" 320x240, template "con fondo"
   on GenerateScreen: SetTag("NombreImagen", 'Gráficos')
   Button "Botón_5" at 278,36 size 26x23; TextOff 'Text'; PictureOff "Gráfico_14"
      on Release: function_efd93a16()
   TextField "Campo de texto_1" at 9,46 size 127x16; Text 'Curvas observables:'
   Button "Botón_1" at 26,73 size 252x25; TextOff 'Temperatura Fermentador'
      on Release: ActivateScreen("Temperatura Fermentador", 0)
   Button "Botón_2" at 26,106 size 252x25; TextOff 'Temperatura Alambique'
      on Release: ActivateScreen("Temperatura Destilador", 0)
   Button "Botón_3" at 26,141 size 252x25; TextOff 'Volumenes del proceso'
      on Release: ActivateScreen("Volumenes", 0)

screen "Configuración" 320x240, template "con fondo"
   on GenerateScreen: SetTag("NombreImagen", 'Configuración')
   GraphicView "Visor de gráficos_1" at 161,55 size 36x30; Picture "Gráfico_18"
      Visibility <- "ModoManualActivado"
   Button "Botón_1" at 19,55 size 136x32; TextOff 'Poner en modo manual'; TextOn 'Poner en modo automatico'; Authorization "Operación"
      on Release: SetBit("ModoManualActivado")
      Visibility <- "ModoManualActivado"
   Button "Botón_2" at 20,142 size 136x32; TextOn 'Poner en modo automatico'; TextOff 'Recetas'; Authorization "Operación"
      on Release: ActivateScreen("Recetas", 0)
   GraphicView "Visor de gráficos_5" at 163,96 size 36x30; Picture "Gráfico_19"
      Visibility <- "ModoManualActivado"
   GraphicView "Visor de gráficos_6" at 161,142 size 36x30; Picture "Gráfico_20"
   Button "Botón_5" at 274,41 size 40x27; TextOff 'Text'; PictureOff "Gráfico_14"
      on Release: function_efd93a16()
   Button "Botón_3" at 20,96 size 136x32; TextOn 'Poner en modo automatico'; TextOff 'Poner en modo automatico'; Authorization "Operación"
      on Release: ResetBit("ModoManualActivado")
      Visibility <- "ModoManualActivado"

screen "Recetas" 320x240, template "con fondo"
   on GenerateScreen: SetTag("NombreImagen", 'Recetas')
   Button "Botón_5" at 274,41 size 40x27; TextOff 'Text'; PictureOff "Gráfico_14"
      on Release: function_efd93a16()
   RecipeView "Visor de recetas_2" at 4,49 size 208x151; Recipe "Whiskey"; Tag4DataRecord "DatosDeRecetas_NombreRecetaActiva"
   TextField "Campo de texto_2" at 218,84 size 96x13; Text 'Estamos haciendo:'
   IOField "Campo ES_1" at 221,109 size 96x23; FormatPattern ????????????????????????????????????????????????????????????????????????????????
      ProcessValue <- "Name"

screen "Temperatura Fermentador" 320x240, template "con fondo"
   on GenerateScreen: SetTag("NombreImagen", 'Gráficos')
   TrendView "Visor de curvas_1" at 7,42 size 299x165

screen "Volumenes" 320x240, template "con fondo"
   on GenerateScreen: SetTag("NombreImagen", 'Gráficos')
   TrendView "Visor de curvas_1" at 9,43 size 302x163

screen "Temperatura Destilador" 320x240, template "con fondo"
   on GenerateScreen: SetTag("NombreImagen", 'Gráficos')
   TrendView "Visor de curvas_1" at 5,43 size 306x163

scheduled task "LeerNombre"
   on Action: function_f41c6f6c("NombreDeUsuario")
*)